(* IEC 61131-3 sources: JingjiangArm/moonboxpro_arm_8.4/Application/Application/任务列表/CommTask/COMM_DIAMONDS/Input_Output (part 3) *)

	i_pstStSysParam^.astStGrpParam_Save[iGrp].rAdjVal_PerTime_Fine			:=	i_pstStParam_Diamonds_WrRd^.arAdjVal_PerTime_Fine[iGrp]   		 	;											(*手动细调调整量*)
	i_pstStSysParam^.astStGrpParam_Save[iGrp].rAdjVal_PerTime_Coarse		:=	i_pstStParam_Diamonds_WrRd^.arAdjVal_PerTime_Coarse[iGrp] 		 	;										(*手动粗调调整量*)
	i_pstStSysParam^.astStGrpParam_Save[iGrp].rVel_HorzdAdj					:=	i_pstStParam_Diamonds_WrRd^.arVel_HorzAdjust[iGrp]        		 	;													(*横向调整速度*)
	i_pstStSysParam^.astStGrpParam_Save[iGrp].rVel_HorzPreRegister			:=	i_pstStParam_Diamonds_WrRd^.arVel_HorzPreRegister[iGrp]   		 	;											(*横向预套准速度*)
	i_pstStSysParam^.astStGrpParam_Save[iGrp].uiNum_If						:=	i_pstStParam_Diamonds_WrRd^.auiNum_If[iGrp]               		 	;														(*放牵减速比-电机侧*)
	i_pstStSysParam^.astStGrpParam_Save[iGrp].uiDen_If						:=	i_pstStParam_Diamonds_WrRd^.auiDen_If[iGrp]               		 	;														(*放牵减速比-传动侧*)
	i_pstStSysParam^.astStGrpParam_Save[iGrp].uiNum_Of						:=	i_pstStParam_Diamonds_WrRd^.auiNum_Of[iGrp]               		 	;														(*收牵减速比-电机侧*)
	i_pstStSysParam^.astStGrpParam_Save[iGrp].uiDen_Of						:=	i_pstStParam_Diamonds_WrRd^.auiDen_Of[iGrp]               		 	;														(*收牵减速比-传动侧*)
	i_pstStSysParam^.astStGrpParam_Save[iGrp].uiNum_Uw						:=	i_pstStParam_Diamonds_WrRd^.auiNum_Uw[iGrp]               		 	;														(*放料减速比-电机侧*)
	i_pstStSysParam^.astStGrpParam_Save[iGrp].uiDen_Uw						:=	i_pstStParam_Diamonds_WrRd^.auiDen_Uw[iGrp]               		 	;														(*放料减速比-传动侧*)
	i_pstStSysParam^.astStGrpParam_Save[iGrp].uiNum_Rw						:=	i_pstStParam_Diamonds_WrRd^.auiNum_Rw[iGrp]               		 	;														(*收料减速比-电机侧*)
	i_pstStSysParam^.astStGrpParam_Save[iGrp].uiDen_Rw						:=	i_pstStParam_Diamonds_WrRd^.auiDen_Rw[iGrp]               		 	;														(*收料减速比-传动侧*)
	i_pstStSysParam^.astStGrpParam_Save[iGrp].uiNum_PrnRoller				:=	i_pstStParam_Diamonds_WrRd^.auiNum_Pu[iGrp]               		 	;												(*色组减速比-电机侧*)
	i_pstStSysParam^.astStGrpParam_Save[iGrp].uiDen_PrnRoller				:=	i_pstStParam_Diamonds_WrRd^.auiDen_Pu[iGrp]               		 	;												(*色组减速比-传动侧*)
	(*待补充-开始|2025.08.07.202603*)
(*	i_pstStSysParam^.astStGrpParam_Save[iGrp].wOutput_IOtestDO_Main[1]		:=	i_pstStParam_Diamonds_WrRd^.awOutput_IOtestDO_Main[iGrp][1]		 	;										(*主面板IO测试输出*)
	i_pstStSysParam^.astStGrpParam_Save[iGrp].wOutput_IOtestDO_Main[2]		:=	i_pstStParam_Diamonds_WrRd^.awOutput_IOtestDO_Main[iGrp][2]		 	;										(*主面板IO测试输出*)
	i_pstStSysParam^.astStGrpParam_Save[iGrp].wOutput_IOtestDO_Main[3]		:=	i_pstStParam_Diamonds_WrRd^.awOutput_IOtestDO_Main[iGrp][3]		 	;										(*主面板IO测试输出*)
	i_pstStSysParam^.astStGrpParam_Save[iGrp].wOutput_IOtestDO_Main[4]		:=	i_pstStParam_Diamonds_WrRd^.awOutput_IOtestDO_Main[iGrp][4]		 	;										(*主面板IO测试输出*)
	i_pstStSysParam^.astStGrpParam_Save[iGrp].wOutput_IOtestDO_Main[5]		:=	i_pstStParam_Diamonds_WrRd^.awOutput_IOtestDO_Main[iGrp][5]		 	;										(*主面板IO测试输出*)
	i_pstStSysParam^.astStGrpParam_Save[iGrp].wOutput_IOtestDO_Main[6]		:=	i_pstStParam_Diamonds_WrRd^.awOutput_IOtestDO_Main[iGrp][6]		 	;										(*主面板IO测试输出*)
	i_pstStSysParam^.astStGrpParam_Save[iGrp].wOutput_IOtestDO_Main[7]		:=	i_pstStParam_Diamonds_WrRd^.awOutput_IOtestDO_Main[iGrp][7]		 	;										(*主面板IO测试输出*)
	i_pstStSysParam^.astStGrpParam_Save[iGrp].wOutput_IOtestDO_Main[8]		:=	i_pstStParam_Diamonds_WrRd^.awOutput_IOtestDO_Main[iGrp][8]		 	;										(*主面板IO测试输出*)

	i_pstStSysParam^.astStGrpParam_Save[iGrp].wOutput_IOtestAO_Main[1]		:=	i_pstStParam_Diamonds_WrRd^.awOutput_IOtestAO_Main[iGrp][1]		 	;									(*主面板IO测试输出*)
	i_pstStSysParam^.astStGrpParam_Save[iGrp].wOutput_IOtestAO_Main[2]		:=	i_pstStParam_Diamonds_WrRd^.awOutput_IOtestAO_Main[iGrp][2]		 	;									(*主面板IO测试输出*)
	i_pstStSysParam^.astStGrpParam_Save[iGrp].wOutput_IOtestAO_Main[3]		:=	i_pstStParam_Diamonds_WrRd^.awOutput_IOtestAO_Main[iGrp][3]		 	;									(*主面板IO测试输出*)
	i_pstStSysParam^.astStGrpParam_Save[iGrp].wOutput_IOtestAO_Main[4]		:=	i_pstStParam_Diamonds_WrRd^.awOutput_IOtestAO_Main[iGrp][4]		 	;									(*主面板IO测试输出*)
	i_pstStSysParam^.astStGrpParam_Save[iGrp].wOutput_IOtestAO_Main[5]		:=	i_pstStParam_Diamonds_WrRd^.awOutput_IOtestAO_Main[iGrp][5]		 	;									(*主面板IO测试输出*)
	i_pstStSysParam^.astStGrpParam_Save[iGrp].wOutput_IOtestAO_Main[6]		:=	i_pstStParam_Diamonds_WrRd^.awOutput_IOtestAO_Main[iGrp][6]		 	;									(*主面板IO测试输出*)
	i_pstStSysParam^.astStGrpParam_Save[iGrp].wOutput_IOtestAO_Main[7]		:=	i_pstStParam_Diamonds_WrRd^.awOutput_IOtestAO_Main[iGrp][7]		 	;									(*主面板IO测试输出*)
	i_pstStSysParam^.astStGrpParam_Save[iGrp].wOutput_IOtestAO_Main[8]		:=	i_pstStParam_Diamonds_WrRd^.awOutput_IOtestAO_Main[iGrp][8]		 	;									(*主面板IO测试输出*)
	i_pstStSysParam^.astStGrpParam_Save[iGrp].wOutput_IOtestAO_Main[9]		:=	i_pstStParam_Diamonds_WrRd^.awOutput_IOtestAO_Main[iGrp][9]		 	;									(*主面板IO测试输出*)
	i_pstStSysParam^.astStGrpParam_Save[iGrp].wOutput_IOtestAO_Main[10]		:=	i_pstStParam_Diamonds_WrRd^.awOutput_IOtestAO_Main[iGrp][10]	 	;										(*主面板IO测试输出*)
	i_pstStSysParam^.astStGrpParam_Save[iGrp].wOutput_IOtestAO_Main[11]		:=	i_pstStParam_Diamonds_WrRd^.awOutput_IOtestAO_Main[iGrp][11]	 	;										(*主面板IO测试输出*)
	i_pstStSysParam^.astStGrpParam_Save[iGrp].wOutput_IOtestAO_Main[12]		:=	i_pstStParam_Diamonds_WrRd^.awOutput_IOtestAO_Main[iGrp][12]	 	;										(*主面板IO测试输出*)
	i_pstStSysParam^.astStGrpParam_Save[iGrp].wOutput_IOtestAO_Main[13]		:=	i_pstStParam_Diamonds_WrRd^.awOutput_IOtestAO_Main[iGrp][13]	 	;										(*主面板IO测试输出*)
	i_pstStSysParam^.astStGrpParam_Save[iGrp].wOutput_IOtestAO_Main[14]		:=	i_pstStParam_Diamonds_WrRd^.awOutput_IOtestAO_Main[iGrp][14]	 	;										(*主面板IO测试输出*)
	i_pstStSysParam^.astStGrpParam_Save[iGrp].wOutput_IOtestAO_Main[15]		:=	i_pstStParam_Diamonds_WrRd^.awOutput_IOtestAO_Main[iGrp][15]	 	;										(*主面板IO测试输出*)
	i_pstStSysParam^.astStGrpParam_Save[iGrp].wOutput_IOtestAO_Main[16]		:=	i_pstStParam_Diamonds_WrRd^.awOutput_IOtestAO_Main[iGrp][16]	 	;										(*主面板IO测试输出*)
*)	(*待补充-结束|2025.08.07.202615*)

	i_pstStSysParam^.astStGrpParam_Save[iGrp].uiPreStopDelayTime_ms		:= 	i_pstStParam_Diamonds_WrRd^.auiPreStopDelayTime_ms[iGrp]    	;
	i_pstStSysParam^.astStGrpParam_Save[iGrp].rVel_Tar_9905				:= 	i_pstStParam_Diamonds_WrRd^.arVel_Tar_9905[iGrp]            	;
	i_pstStSysParam^.astStGrpParam_UnSave[iGrp].iAxisId_StepTest_V		:= 	i_pstStParam_Diamonds_WrRd^.aiAxisId_StepTest_V[iGrp]       	;
	i_pstStSysParam^.astStGrpParam_UnSave[iGrp].iInterval_StepTest12		:= 	i_pstStParam_Diamonds_WrRd^.aiInterval_StepTest12[iGrp]     	;
	i_pstStSysParam^.astStGrpParam_Save[iGrp].iMicron_StepTest1_V		:= 	i_pstStParam_Diamonds_WrRd^.aiMicron_StepTest1_V[iGrp]      	;
	i_pstStSysParam^.astStGrpParam_Save[iGrp].iMicron_StepTest2_V		:= 	i_pstStParam_Diamonds_WrRd^.aiMicron_StepTest2_V[iGrp]      	;
	i_pstStSysParam^.astStGrpParam_Save[iGrp].byKalmanFilterType_Rw		:= 	i_pstStParam_Diamonds_WrRd^.abyKalmanFilterType_Rw[iGrp]    	;
	IF i_pstStParam_Diamonds_WrRd^.abyStructParanInitEn_Rw[iGrp]<>0 THEN
		i_pstStSysParam^.astStGrpParam_Save[iGrp].byStructParanInitEn_Rw 	:= 	i_pstStParam_Diamonds_WrRd^.abyStructParanInitEn_Rw[iGrp]   	;
	END_IF
	i_pstStSysParam^.astStGrpParam_Save[iGrp].rR_K_MinBeat_Rw	    	:= 	i_pstStParam_Diamonds_WrRd^.arR_K_MinBeat_Rw[iGrp]          	;
	i_pstStSysParam^.astStGrpParam_Save[iGrp].iN_MinBeat_Rw	        	:= 	i_pstStParam_Diamonds_WrRd^.aiN_MinBeat_Rw[iGrp]            	;
	i_pstStSysParam^.astStGrpParam_Save[iGrp].rR_K_LQR_Rw	        	:= 	i_pstStParam_Diamonds_WrRd^.arR_K_LQR_Rw[iGrp]              	;

	i_pstStSysParam^.astStGrpParam_Save[iGrp].rN_LQR_Rw	            		:= i_pstStParam_Diamonds_WrRd^.arN_LQR_Rw[iGrp]	               		;
	i_pstStSysParam^.astStGrpParam_Save[iGrp].rKc_Rw	            		:= i_pstStParam_Diamonds_WrRd^.arKc_Rw[iGrp]	                   	;
	i_pstStSysParam^.astStGrpParam_Save[iGrp].rKc_Rw_AccDec	        		:= i_pstStParam_Diamonds_WrRd^.arKc_Rw_AccDec[iGrp]	           		;
	i_pstStSysParam^.astStGrpParam_Save[iGrp].rWc_LowPass_Diam_Rw			:= i_pstStParam_Diamonds_WrRd^.arWc_LowPass_Diam_Rw[iGrp]	   		;
	i_pstStSysParam^.astStGrpParam_Save[iGrp].byKalmanFilterType_Uw 		:= i_pstStParam_Diamonds_WrRd^.abyKalmanFilterType_Uw[iGrp] 	   	;
	IF i_pstStParam_Diamonds_WrRd^.abyStructParanInitEn_Uw[iGrp]<>0 THEN
		i_pstStSysParam^.astStGrpParam_Save[iGrp].byStructParanInitEn_Uw		:= i_pstStParam_Diamonds_WrRd^.abyStructParanInitEn_Uw[iGrp]	   	;
	END_IF
	SysMemCpy(
		ADR(i_pstStSysParam^.astStGrpParam_Save[iGrp].stModelParam_Uw),
		ADR(i_pstStParam_Diamonds_WrRd^.astModelParam_Uw[iGrp]),
		SIZEOF(i_pstStSysParam^.astStGrpParam_Save[iGrp].stModelParam_Uw));
	SysMemCpy(
		ADR(i_pstStSysParam^.astStGrpParam_Save[iGrp].stInvariant_Parameters_Uw),
		ADR(i_pstStParam_Diamonds_WrRd^.astInvariant_Parameters_Uw[iGrp]),
		SIZEOF(i_pstStSysParam^.astStGrpParam_Save[iGrp].stInvariant_Parameters_Uw));
	SysMemCpy(
		ADR(i_pstStSysParam^.astStGrpParam_Save[iGrp].stPI_Parameters_Uw),
		ADR(i_pstStParam_Diamonds_WrRd^.astPI_Parameters_Uw[iGrp]),
		SIZEOF(i_pstStSysParam^.astStGrpParam_Save[iGrp].stPI_Parameters_Uw));
	SysMemCpy(
		ADR(i_pstStSysParam^.astStGrpParam_Save[iGrp].stPI_Parameters_Uw_AccDec),
		ADR(i_pstStParam_Diamonds_WrRd^.astPI_Parameters_Uw_AccDec[iGrp]),
		SIZEOF(i_pstStSysParam^.astStGrpParam_Save[iGrp].stPI_Parameters_Uw_AccDec));

	SysMemCpy(
		ADR(i_pstStSysParam^.astStGrpParam_Save[iGrp].stModelParam_Rw),
		ADR(i_pstStParam_Diamonds_WrRd^.astModelParam_Rw[iGrp]),
		SIZEOF(i_pstStSysParam^.astStGrpParam_Save[iGrp].stModelParam_Rw));
	SysMemCpy(
		ADR(i_pstStSysParam^.astStGrpParam_Save[iGrp].stInvariant_Parameters_Rw),
		ADR(i_pstStParam_Diamonds_WrRd^.astInvariant_Parameters_Rw[iGrp]),
		SIZEOF(i_pstStSysParam^.astStGrpParam_Save[iGrp].stInvariant_Parameters_Rw));
	SysMemCpy(
		ADR(i_pstStSysParam^.astStGrpParam_Save[iGrp].stPI_Parameters_Rw),
		ADR(i_pstStParam_Diamonds_WrRd^.astPI_Parameters_Rw[iGrp]),
		SIZEOF(i_pstStSysParam^.astStGrpParam_Save[iGrp].stPI_Parameters_Rw));
	SysMemCpy(
		ADR(i_pstStSysParam^.astStGrpParam_Save[iGrp].stPI_Parameters_Rw_AccDec),
		ADR(i_pstStParam_Diamonds_WrRd^.astPI_Parameters_Rw_AccDec[iGrp]),
		SIZEOF(i_pstStSysParam^.astStGrpParam_Save[iGrp].stPI_Parameters_Rw_AccDec));

	i_pstStSysParam^.astStGrpParam_Save[iGrp].rR_K_MinBeat_Uw    			:= i_pstStParam_Diamonds_WrRd^.arR_K_MinBeat_Uw[iGrp]    			;
	i_pstStSysParam^.astStGrpParam_Save[iGrp].iN_MinBeat_Uw      			:= i_pstStParam_Diamonds_WrRd^.aiN_MinBeat_Uw[iGrp]      			;
	i_pstStSysParam^.astStGrpParam_Save[iGrp].rR_K_LQR_Uw        			:= i_pstStParam_Diamonds_WrRd^.arR_K_LQR_Uw[iGrp]        			;
	i_pstStSysParam^.astStGrpParam_Save[iGrp].rN_LQR_Uw          			:= i_pstStParam_Diamonds_WrRd^.arN_LQR_Uw[iGrp]          			;
	i_pstStSysParam^.astStGrpParam_Save[iGrp].rKc_Uw             			:= i_pstStParam_Diamonds_WrRd^.arKc_Uw[iGrp]             			;
	i_pstStSysParam^.astStGrpParam_Save[iGrp].rKc_Uw_AccDec      			:= i_pstStParam_Diamonds_WrRd^.arKc_Uw_AccDec[iGrp]      			;
	i_pstStSysParam^.astStGrpParam_Save[iGrp].rWc_LowPass_Diam_Uw			:= i_pstStParam_Diamonds_WrRd^.arWc_LowPass_Diam_Uw[iGrp]			;

	i_pstStSysParam^.astStGrpParam_Save[iGrp].rWn_Uw         				:= i_pstStParam_Diamonds_WrRd^.arWn_Uw[iGrp]         	      		;
	i_pstStSysParam^.astStGrpParam_Save[iGrp].rBw_Uw         				:= i_pstStParam_Diamonds_WrRd^.arBw_Uw[iGrp]         	      		;
	i_pstStSysParam^.astStGrpParam_Save[iGrp].rDp_Uw         				:= i_pstStParam_Diamonds_WrRd^.arDp_Uw[iGrp]         	      		;
	i_pstStSysParam^.astStGrpParam_Save[iGrp].iWorkMode_Pid					:= i_pstStParam_Diamonds_WrRd^.aiWorkMode_Pid[iGrp]		  			;
	i_pstStSysParam^.astStGrpParam_Save[iGrp].rFilmLenth_InUnit  			:= i_pstStParam_Diamonds_WrRd^.arFilmLenth_InUnit[iGrp]	   			;

	(*增加裁切时间集处理2025.9.11.193948*)
	//2026.05.20.214715 替换为直接赋值 by liu.yt
	i_pstStSysParam^.astStGrpParam_UnSave[iGrp].stStTimeSet_DnCut_UpCut_Uw_Hmi:=i_pstStParam_Diamonds_WrRd^.astStTimeSet_DnCut_UpCut_Uw_Hmi[iGrp];
	//2026.05.21.085510 补充收料
	i_pstStSysParam^.astStGrpParam_UnSave[iGrp].stStTimeSet_DnCut_UpCut_RW_Hmi:=i_pstStParam_Diamonds_WrRd^.astStTimeSet_DnCut_UpCut_Rw_Hmi[iGrp];

	i_pstStSysParam^.astStGrpParam_Save[iGrp].byAIType_Uw:= i_pstStParam_Diamonds_WrRd^.abyAIType_Uw[iGrp];
	i_pstStSysParam^.astStGrpParam_Save[iGrp].byAIType_Rw:= i_pstStParam_Diamonds_WrRd^.abyAIType_Rw[iGrp];
	i_pstStSysParam^.astStGrpParam_Save[iGrp].byAIType_If:= i_pstStParam_Diamonds_WrRd^.abyAIType_If[iGrp];
	i_pstStSysParam^.astStGrpParam_Save[iGrp].byAIType_Of:= i_pstStParam_Diamonds_WrRd^.abyAIType_Of[iGrp];
(*2025.10.24.134439||增加变量*)
	i_pstStSysParam^.astStGrpParam_Save[iGrp].byAlarmHold_PreCut_Uw:= i_pstStParam_Diamonds_WrRd^.abyAlarmHold_PreCut_Uw[iGrp];
	i_pstStSysParam^.astStGrpParam_Save[iGrp].byFilmType:= i_pstStParam_Diamonds_WrRd^.abyFilmType[iGrp];
	i_pstStSysParam^.astStGrpParam_Save[iGrp].uiUseTime_Diam_Min_Uw:= i_pstStParam_Diamonds_WrRd^.auiUseTime_Diam_Min_Uw[iGrp];
	i_pstStSysParam^.astStGrpParam_Save[iGrp].uiUseTime_Diam_Min_Rw:= i_pstStParam_Diamonds_WrRd^.auiUseTime_Diam_Min_Rw[iGrp];

(*2025.11.5.154653*)
	i_pstStSysParam^.astStGrpParam_Save[iGrp].iUpperFreq_InkRoller:= i_pstStParam_Diamonds_WrRd^.aiUpperFreq_InkRoller[iGrp];
	i_pstStSysParam^.astStGrpParam_Save[iGrp].iVelSa_InkRollerRun:= i_pstStParam_Diamonds_WrRd^.aiVelSa_InkRollerRun[iGrp];
	i_pstStSysParam^.astStGrpParam_Save[iGrp].iFrq_InkRollerMin:= i_pstStParam_Diamonds_WrRd^.aiFrq_InkRollerMin[iGrp];
	i_pstStSysParam^.astStGrpParam_Save[iGrp].iFrq_InkRollerMax:= i_pstStParam_Diamonds_WrRd^.aiFrq_InkRollerMax[iGrp];
	i_pstStSysParam^.astStGrpParam_Save[iGrp].iVel_InkRollerMin:= i_pstStParam_Diamonds_WrRd^.aiVel_InkRollerMin[iGrp];
	i_pstStSysParam^.astStGrpParam_Save[iGrp].iVel_InkRollerMax:= i_pstStParam_Diamonds_WrRd^.aiVel_InkRollerMax[iGrp];
	i_pstStSysParam^.astStGrpParam_UnSave[iGrp].byPseudoRandomId:= i_pstStParam_Diamonds_WrRd^.abyPseudoRandomId[iGrp];
	i_pstStSysParam^.astStGrpParam_Save[iGrp].rHz_PreHotAir_ManuallySet:= i_pstStParam_Diamonds_WrRd^.arHz_PreHotAir_ManuallySet[iGrp];
	i_pstStSysParam^.astStGrpParam_Save[iGrp].rSV_PreHeating:= i_pstStParam_Diamonds_WrRd^.arSV_PreHeating[iGrp];
	i_pstStSysParam^.astStGrpParam_Save[iGrp].rHz_Scraper_ManuallySet:= i_pstStParam_Diamonds_WrRd^.arHz_Scraper_ManuallySet[iGrp];
	i_pstStSysParam^.astStGrpParam_Save[iGrp].rCoeff_Scraper_Auto:= i_pstStParam_Diamonds_WrRd^.arCoeff_Scraper_Auto[iGrp];
	i_pstStSysParam^.astStGrpParam_Save[iGrp].rHz_InkRoller_ManuallySet:= i_pstStParam_Diamonds_WrRd^.arHz_InkRoller_ManuallySet[iGrp];
	i_pstStSysParam^.astStGrpParam_Save[iGrp].rCoeff_InkRoller:= i_pstStParam_Diamonds_WrRd^.arCoeff_InkRoller_Auto[iGrp];
//2026.1.6.095943增加一些变量
	i_pstStSysParam^.astStGrpParam_Save[iGrp].rLength_Band_Confirm:= i_pstStParam_Diamonds_WrRd^.arLength_Band_Confirm[iGrp];
	i_pstStSysParam^.astStGrpParam_Save[iGrp].rPressure_Tar:= i_pstStParam_Diamonds_WrRd^.arPressure_Tar[iGrp];
// 	xSwitch_TensionAdjust_QH					: BIT;
// 	xSwitch_PrnLenAdj_Follow_QH					: BIT;
	i_pstStSysParam^.stStSysParam_Save.dwCtlSwitchRef.3:= i_pstStParam_Diamonds_WrRd^.astBitStWrRd_Switch_Grp[iGrp].xSwitch_TensionAdjust_QH;
	i_pstStSysParam^.stStSysParam_Save.dwCtlSwitchRef.2:= i_pstStParam_Diamonds_WrRd^.astBitStWrRd_Switch_Grp[iGrp].xSwitch_PrnLenAdj_Follow_QH;

	//2026.2.2.165944||新增界面的一些内容|Niu/j
	i_pstStSysParam^.astStGrpParam_Save[iGrp].rScrewPitch_PrnRoller_Pressure:=
					i_pstStParam_Diamonds_WrRd^.arScrewPitch_PrnRoller_Pressure[iGrp];
	i_pstStSysParam^.astStGrpParam_Save[iGrp].uiNum_PrnRoller_Pressure:=
					i_pstStParam_Diamonds_WrRd^.auiNum_PrnRoller_Pressure[iGrp];
	i_pstStSysParam^.astStGrpParam_Save[iGrp].uiDen_PrnRoller_Pressure:=
					i_pstStParam_Diamonds_WrRd^.auiDen_PrnRoller_Pressure[iGrp];

	i_pstStSysParam^.astStGrpParam_Save[iGrp].rScrewPitch_NetRoller_Pressure:=
					i_pstStParam_Diamonds_WrRd^.arScrewPitch_NetRoller_Pressure[iGrp];
	i_pstStSysParam^.astStGrpParam_Save[iGrp].uiNum_NetRoller_Pressure:=
					i_pstStParam_Diamonds_WrRd^.auiNum_NetRoller_Pressure[iGrp];
	i_pstStSysParam^.astStGrpParam_Save[iGrp].uiDen_NetRoller_Pressure:=
					i_pstStParam_Diamonds_WrRd^.auiDen_NetRoller_Pressure[iGrp];

	i_pstStSysParam^.astStGrpParam_Save[iGrp].rScrewPitch_StrRoller_Pressure:=
					i_pstStParam_Diamonds_WrRd^.arScrewPitch_StrRoller_Pressure[iGrp];
	i_pstStSysParam^.astStGrpParam_Save[iGrp].uiNum_StrRoller_Pressure:=
					i_pstStParam_Diamonds_WrRd^.auiNum_StrRoller_Pressure[iGrp];
	i_pstStSysParam^.astStGrpParam_Save[iGrp].uiDen_StrRoller_Pressure:=
					i_pstStParam_Diamonds_WrRd^.auiDen_StrRoller_Pressure[iGrp];

	i_pstStSysParam^.astStGrpParam_Save[iGrp].rScrewPitch_Horz:=
					i_pstStParam_Diamonds_WrRd^.arScrewPitch_Horz[iGrp];
	i_pstStSysParam^.astStGrpParam_Save[iGrp].uiNum_Horz:=
					i_pstStParam_Diamonds_WrRd^.auiNum_Horz[iGrp];
	i_pstStSysParam^.astStGrpParam_Save[iGrp].uiDen_Horz:=
					i_pstStParam_Diamonds_WrRd^.auiDen_Horz[iGrp];

	i_pstStSysParam^.astStRSV_GrpParam_Save[iGrp].rVel_UVstartVel:= i_pstStParam_Diamonds_WrRd^.arVel_UVstartVel[iGrp];

	//2026.02.28.144731 | + | 上下裁切换
	i_pstStSysParam^.astStGrpParam_Save[iGrp].xSwitch_Change_CutterOnTop_HMI_Uw:=i_pstStParam_Diamonds_WrRd^.astBitStWrRd_Switch_Grp[iGrp].xSwitch_Change_CutterOnTop_HMI_Uw;(*上下裁切换*)
	i_pstStSysParam^.astStGrpParam_Save[iGrp].xSwitch_Change_CutterOnTop_HMI_Rw:=i_pstStParam_Diamonds_WrRd^.astBitStWrRd_Switch_Grp[iGrp].xSwitch_Change_CutterOnTop_HMI_Rw;(*上下裁切换*)

	//2026.03.11.100402 | + | 使用Bit22作为压力电机自动合压开关
	i_pstStSysParam^.astStGrpParam_Save[iGrp].wCtl_Pressure_Up_Dn.0:=i_pstStParam_Diamonds_WrRd^.astBitStWrRd_Switch_Grp[iGrp].xSwitch_PressureAuto_Up_Dn;

	//2026.03.11.114928 | + | 使用Bit24作为停机维持使能的开关
	i_pstStSysParam^.astStGrpParam_Save[iGrp].dwExtBitCtlFlag.21 :=i_pstStParam_Diamonds_WrRd^.astBitStWrRd_Switch_Grp[iGrp].xSwitch_KeepServoOn;

	//2026.02.25.100358 | + | 使用Bit23作为控制天枢存储数据的开关
	i_pstStSysParam^.astStGrpParam_Save[iGrp].dwExtBitCtlFlag.22 :=i_pstStParam_Diamonds_WrRd^.astBitStWrRd_Switch_Grp[iGrp].xSwitch_SaveData_GNS;

	//2026.03.27.175514 | + | 给超旭同步秦华的金刚清除报警功能    2026.1.27.141112 | + | 增加清除报警的功能
	IF 	i_pstStParam_Diamonds_WrRd^.astBitStWrRd_Switch_Grp[iGrp].xSwitch_ClearSysAlarm THEN
		i_pstStParam_Diamonds_WrRd^.astBitStWrRd_Switch_Grp[iGrp].xSwitch_ClearSysAlarm := FALSE;
		g_xClrAlr_HMI := TRUE;
	END_IF
	//2026.04.01.165429 增加总匀墨 Hou.N
	i_pstStSysParam^.astStRSV_GrpParam_UnSave[iGrp].xSwitch_GrpInkEn :=i_pstStParam_Diamonds_WrRd^.astBitStWrRd_Switch_Grp[iGrp].xSwitch_GrpInkEn;
	IF i_pstStParam_Diamonds_WrRd^.astBitStWrRd_Switch_Grp[iGrp].xBtn_ChangeFilmDn_Uw THEN
		i_pstStSysParam^.astStGrpParam_UnSave[iGrp].xCurAxisDia_Uw_Wr:= i_pstStParam_Diamonds_WrRd^.astBitStWrRd_Switch_Grp[iGrp].xBtn_ChangeFilmDn_Uw;
		i_pstStParam_Diamonds_WrRd^.astBitStWrRd_Switch_Grp[iGrp].xBtn_ChangeFilmDn_Uw:= FALSE;
	END_IF
	IF i_pstStParam_Diamonds_WrRd^.astBitStWrRd_Switch_Grp[iGrp].xBtn_ChangeFilmDn_Rw THEN
		i_pstStSysParam^.astStGrpParam_UnSave[iGrp].xCurAxisDia_Rw_Wr:= i_pstStParam_Diamonds_WrRd^.astBitStWrRd_Switch_Grp[iGrp].xBtn_ChangeFilmDn_Rw;
		i_pstStParam_Diamonds_WrRd^.astBitStWrRd_Switch_Grp[iGrp].xBtn_ChangeFilmDn_Rw:= FALSE;
	END_IF
//2026.5.9.172241
	//增加全自动套印相关变量的通讯；2026.4.6.112942|niu.j
	i_pstStSysParam^.astStRSV_GrpParam_UnSave[iGrp].xStartAutoFind:=
		i_pstStParam_Diamonds_WrRd^.astBitStWrRd_Switch_Grp[iGrp].xSwitch_StartAutoFind;
//2026.04.06.141649最终需要放开
	i_pstStSysParam^.astStRSV_GrpParam_Save[iGrp].xSwitch_EnFastPress:=
		i_pstStParam_Diamonds_WrRd^.astBitStWrRd_Switch_Grp[iGrp].xSwitch_EnFastPress;
	i_pstStSysParam^.astStRSV_GrpParam_UnSave[iGrp].xSwitch_SaveRS2file:=
		i_pstStParam_Diamonds_WrRd^.astBitStWrRd_Switch_Grp[iGrp].xSwitch_SaveRS2file;
	i_pstStSysParam^.astStRSV_GrpParam_UnSave[iGrp].xSwitch_RFailure:=
		i_pstStParam_Diamonds_WrRd^.astBitStWrRd_Switch_Grp[iGrp].xSwitch_RFailure;
	i_pstStSysParam^.astStRSV_GrpParam_UnSave[iGrp].xSwitch_FFailure:=
		i_pstStParam_Diamonds_WrRd^.astBitStWrRd_Switch_Grp[iGrp].xSwitch_FFailure;
	i_pstStSysParam^.astStRSV_GrpParam_Save[iGrp].rWidth_Mark_Max:=
			i_pstStParam_Diamonds_WrRd^.arWidth_Mark_Max[iGrp];
	i_pstStSysParam^.astStRSV_GrpParam_Save[iGrp].rWidth_Mark_Min:=
			i_pstStParam_Diamonds_WrRd^.arWidth_Mark_Min[iGrp];
	i_pstStSysParam^.astStRSV_GrpParam_Save[iGrp].rMaxGap:=
			i_pstStParam_Diamonds_WrRd^.arMaxGap[iGrp];
	i_pstStSysParam^.astStRSV_GrpParam_Save[iGrp].bySimilarityThreshold:=
			REAL_TO_BYTE(i_pstStParam_Diamonds_WrRd^.arSimilarityThreshold[iGrp]);
	i_pstStSysParam^.astStRSV_GrpParam_Save[iGrp].byMeanOffset:=
			i_pstStParam_Diamonds_WrRd^.abyMeanOffset[iGrp];
	i_pstStSysParam^.astStRSV_GrpParam_Save[iGrp].bySignalType:=
			i_pstStParam_Diamonds_WrRd^.abySignalType[iGrp];
	i_pstStSysParam^.astStRSV_GrpParam_Save[iGrp].rOuterCoff:=
			i_pstStParam_Diamonds_WrRd^.arOuterCoff[iGrp];
	i_pstStSysParam^.astStRSV_GrpParam_Save[iGrp].rInnerCoff:=
			i_pstStParam_Diamonds_WrRd^.arInnerCoff[iGrp];
	FOR iN:=1 TO 15 BY 1 DO
		IF iN<=2 THEN
			i_pstStSysParam^.astStRSV_GrpParam_Save[iGrp].arFiberMove[iN]:=
						i_pstStParam_Diamonds_WrRd^.arFiberMove[iGrp,iN];
		END_IF
		i_pstStSysParam^.astStRSV_GrpParam_Save[iGrp].arModeMsg[iN]:=
					i_pstStParam_Diamonds_WrRd^.arModeMsg[iGrp,iN];
	END_FOR

	//2026.04.10.110541 增加伪随机pid按钮处理
	i_pstStSysParam^.astStGrpParam_UnSave[iGrp].bySetTestPid_Uw:=i_pstStParam_Diamonds_WrRd^.abySetTestPid_Uw[iGrp];

//2026.4.10.092048增加界面计米清零计数
	IF abyPreCount_ClrPrn[iGrp,1]= i_pstStSysParam^.astStGrpParam_UnSave[iGrp].abyClrPrnLenCount_Rw[1] THEN
		i_pstStSysParam^.astStGrpParam_UnSave[iGrp].abyClrPrnLenCount_Rw[1]:= i_pstStParam_Diamonds_WrRd^.abyClrPrnLenCount[iGrp,1];
	END_IF
	abyPreCount_ClrPrn[iGrp,1]:= i_pstStSysParam^.astStGrpParam_UnSave[iGrp].abyClrPrnLenCount_Rw[1];

	IF abyPreCount_ClrPrn[iGrp,2]= i_pstStSysParam^.astStGrpParam_UnSave[iGrp].abyClrPrnLenCount_Rw[2] THEN
		i_pstStSysParam^.astStGrpParam_UnSave[iGrp].abyClrPrnLenCount_Rw[2]:= i_pstStParam_Diamonds_WrRd^.abyClrPrnLenCount[iGrp,2];
	END_IF
	abyPreCount_ClrPrn[iGrp,2]:= i_pstStSysParam^.astStGrpParam_UnSave[iGrp].abyClrPrnLenCount_Rw[2];

	IF abyPreCount_ClrPrn[iGrp,3]= i_pstStSysParam^.astStGrpParam_UnSave[iGrp].abyClrPrnLenCount_Rw[3] THEN
		i_pstStSysParam^.astStGrpParam_UnSave[iGrp].abyClrPrnLenCount_Rw[3]:= i_pstStParam_Diamonds_WrRd^.abyClrPrnLenCount[iGrp,3];
	END_IF
	abyPreCount_ClrPrn[iGrp,3]:= i_pstStSysParam^.astStGrpParam_UnSave[iGrp].abyClrPrnLenCount_Rw[3];
//增加完成2026.4.10.092101

//2026.5.12.161016增加速度规划方式的通讯
	i_pstStSysParam^.astStGrpParam_Save[iGrp].byAutoAccDecCurve:= i_pstStParam_Diamonds_WrRd^.abyAutoAccDecCurve[iGrp];
	//2026.05.14.151130 新增自动停机、网辊离压速度
    i_pstStSysParam^.astStRSV_GrpParam_Save[iGrp].rRemainDia_stop := i_pstStParam_Diamonds_WrRd^.arRemainDia_stop[iGrp];
    i_pstStSysParam^.astStRSV_GrpParam_Save[iGrp].rMaxErr_GantryTrap := i_pstStParam_Diamonds_WrRd^.arMaxErr_GantryTrap[iGrp];
    i_pstStSysParam^.astStGrpParam_Save[iGrp].rVel_NetReturn := i_pstStParam_Diamonds_WrRd^.arVel_NetReturn[iGrp];
   	i_pstStSysParam^.astStRSV_GrpParam_Save[iGrp].xIsAutoStop :=i_pstStParam_Diamonds_WrRd^.astBitStWrRd_Switch_Grp[iGrp].xSwitch_En_AutoStop;
	//2026.05.15.85606 新增电晕启动速度
	i_pstStSysParam^.astStRSV_GrpParam_Save[iGrp].rVel_CoronaVel:= i_pstStParam_Diamonds_WrRd^.arVel_CoronaVel[iGrp];
	(*2026.05.26.155252+*)
	i_pstStSysParam^.astStGrpParam_UnSave[iGrp].xAutoAccDec_Hmi:=i_pstStParam_Diamonds_WrRd^.astBitStWrRd_Switch_Grp[iGrp].xAutoAccDec_Hmi;

	//2026.05.24.135821 光纤行走部分
	i_pstStSysParam^.astStRSV_GrpParam_Save[iGrp].iFiberMoveVel:=i_pstStParam_Diamonds_WrRd^.aiFiberMoveVel[iGrp];
	i_pstStSysParam^.astStRSV_GrpParam_UnSave[iGrp].rFiberMoveDistance_AllUnit:=i_pstStParam_Diamonds_WrRd^.arFiberMoveDistance_AllUnit[iGrp];
	i_pstStSysParam^.astStRSV_GrpParam_Save[iGrp].byFiberMove_MicroMoveStep:=i_pstStParam_Diamonds_WrRd^.abyFiberMove_MicroMoveStep[iGrp];
	i_pstStSysParam^.astStRSV_GrpParam_UnSave[iGrp].xFiberMove_DebugMode :=i_pstStParam_Diamonds_WrRd^.astBitStWrRd_Switch_Grp[iGrp].xFiberMove_DebugMode;
	i_pstStSysParam^.astStRSV_GrpParam_UnSave[iGrp].xFiberMoveDisRunStart_AllUnit :=i_pstStParam_Diamonds_WrRd^.astBitStWrRd_Switch_Grp[iGrp].xFiberMoveDisRunStart_AllUnit;
	i_pstStSysParam^.astStRSV_GrpParam_Save[iGrp].xUseOnline_FiberMove :=i_pstStParam_Diamonds_WrRd^.astBitStWrRd_Switch_Grp[iGrp].xUseOnline_FiberMove;
	i_pstStSysParam^.astStRSV_GrpParam_UnSave[iGrp].xFiberMoveConfirm_AllUnit :=i_pstStParam_Diamonds_WrRd^.astBitStWrRd_Switch_Grp[iGrp].xFiberMoveConfirm_AllUnit;
	i_pstStSysParam^.astStRSV_GrpParam_UnSave[iGrp].xFiberMovePosCal_ByUnit :=i_pstStParam_Diamonds_WrRd^.astBitStWrRd_Switch_Grp[iGrp].xFiberMovePosCal_ByUnit;
	i_pstStSysParam^.astStRSV_GrpParam_UnSave[iGrp].xFiberMovePosCal_ByOnline :=i_pstStParam_Diamonds_WrRd^.astBitStWrRd_Switch_Grp[iGrp].xFiberMovePosCal_ByOnline;
	i_pstStSysParam^.astStRSV_GrpParam_Save[iGrp].xFiberMove_Negative_AdjustByUnit :=i_pstStParam_Diamonds_WrRd^.astBitStWrRd_Switch_Grp[iGrp].xFiberMove_Negative_AdjustByUnit;
	i_pstStSysParam^.astStRSV_GrpParam_Save[iGrp].xFiberMove_Negative_AdjustByOnline :=i_pstStParam_Diamonds_WrRd^.astBitStWrRd_Switch_Grp[iGrp].xFiberMove_Negative_AdjustByOnline;

//2026.5.15.112026增加卷径检测变量输入
	FOR iK:=1 TO 4 BY 1 DO
		IF arStdVol_Coef_Axis_Hmi_Bak[iGrp,iK]= i_pstStSysParam^.astStGrpParam_UnSave[iGrp].alrStdVol_Coef_Axis_Hmi[iK] THEN
			i_pstStSysParam^.astStGrpParam_UnSave[iGrp].alrStdVol_Coef_Axis_Hmi[iK]:= i_pstStParam_Diamonds_WrRd^.arStdVol_Coef_Axis_Hmi[iGrp,iK];
		END_IF
		arStdVol_Coef_Axis_Hmi_Bak[iGrp,iK]:= i_pstStSysParam^.astStGrpParam_UnSave[iGrp].alrStdVol_Coef_Axis_Hmi[iK];
		IF arStdVol_Diam_Axis_Hmi_Bak[iGrp,iK]= i_pstStSysParam^.astStGrpParam_UnSave[iGrp].alrStdVol_Diam_Axis_Hmi[iK] THEN
			i_pstStSysParam^.astStGrpParam_UnSave[iGrp].alrStdVol_Diam_Axis_Hmi[iK]:=i_pstStParam_Diamonds_WrRd^.arStdVol_Diam_Axis_Hmi[iGrp,iK];
		END_IF
		arStdVol_Diam_Axis_Hmi_Bak[iGrp,iK]:= i_pstStSysParam^.astStGrpParam_UnSave[iGrp].alrStdVol_Diam_Axis_Hmi[iK];
		IF arStdVol_Volt_Axis_Hmi_Bak[iGrp,iK]= i_pstStSysParam^.astStGrpParam_UnSave[iGrp].alrStdVol_Volt_Axis_Hmi[iK] THEN
			i_pstStSysParam^.astStGrpParam_UnSave[iGrp].alrStdVol_Volt_Axis_Hmi[iK]:= i_pstStParam_Diamonds_WrRd^.arStdVol_Volt_Axis_Hmi[iGrp,iK];
		END_IF
		arStdVol_Volt_Axis_Hmi_Bak[iGrp,iK]:= i_pstStSysParam^.astStGrpParam_UnSave[iGrp].alrStdVol_Volt_Axis_Hmi[iK];
	END_FOR
	IF arStdVol_Coef_Axis_Hmi_Bak[iGrp,0]= i_pstStSysParam^.astStGrpParam_UnSave[iGrp].alrStdVol_Coef_Axis_Hmi[0] THEN
		i_pstStSysParam^.astStGrpParam_UnSave[iGrp].alrStdVol_Coef_Axis_Hmi[0]:= i_pstStParam_Diamonds_WrRd^.arStdVol_Coef_Axis_Hmi[iGrp,0];
	END_IF
	arStdVol_Coef_Axis_Hmi_Bak[iGrp,0]:= i_pstStSysParam^.astStGrpParam_UnSave[iGrp].alrStdVol_Coef_Axis_Hmi[0];
END_FOR
(*轴参数|2025.08.07.101610*)
FOR iUnitId:= 1 TO MAX_UNIT_NUM BY 1 DO
	//2026.04.03.115045
	IF axSwitch_AutoAdjust_V_Unit[iUnitId]= i_pstStSysParam^.astStUnitParam_Save[iUnitId].dwFlag_Sts.0 THEN
		i_pstStSysParam^.astStUnitParam_Save[iUnitId].dwFlag_Sts.0 	:=		i_pstStParam_Diamonds_WrRd^.astStWrRd_UnitParam[iUnitId].stBitStWrRd_Switch_Unit.xSwitch_AutoAdjust_V_Unit			 ;			(*整机纵向自动调整开关*)
	END_IF
	axSwitch_AutoAdjust_V_Unit[iUnitId]:= i_pstStSysParam^.astStUnitParam_Save[iUnitId].dwFlag_Sts.0;
	i_pstStSysParam^.astStUnitParam_Save[iUnitId].dwFlag_Sts.1 	:=		i_pstStParam_Diamonds_WrRd^.astStWrRd_UnitParam[iUnitId].stBitStWrRd_Switch_Unit.xSwitch_AutoAdjust_H_Unit			 ;			(*整机纵向自动调整开关*)
	i_pstStSysParam^.astStUnitParam_Save[iUnitId].xEnable_arc 	:=		i_pstStParam_Diamonds_WrRd^.astStWrRd_UnitParam[iUnitId].stBitStWrRd_Switch_Unit.xSwitch_ThisUnitEna ;			(*色组套印开关*)
	i_pstStSysParam^.astStUnitParam_Save[iUnitId].dwFlag_Ctl.0:= i_pstStParam_Diamonds_WrRd^.astStWrRd_UnitParam[iUnitId].stBitStWrRd_Switch_Unit.xSwitch_Horz ;(*横向开关*)
	i_pstStSysParam^.astStUnitParam_Save[iUnitId].dwFlag_Ctl.1:= i_pstStParam_Diamonds_WrRd^.astStWrRd_UnitParam[iUnitId].stBitStWrRd_Switch_Unit.xSwitch_DoorBaseLn	 ;(*门内基线开关*)
	i_pstStSysParam^.astStUnitParam_Save[iUnitId].dwFlag_Ctl.4:= i_pstStParam_Diamonds_WrRd^.astStWrRd_UnitParam[iUnitId].stBitStWrRd_Switch_Unit.xSwitch_AdjRev_V ;(*横向调整反*)
	i_pstStSysParam^.astStUnitParam_Save[iUnitId].dwFlag_Ctl.5:= i_pstStParam_Diamonds_WrRd^.astStWrRd_UnitParam[iUnitId].stBitStWrRd_Switch_Unit.xSwitch_AdjRev_H ;(*横向调整反*)
	i_pstStSysParam^.astStUnitParam_Save[iUnitId].byCouplingMask.2:= i_pstStParam_Diamonds_WrRd^.astStWrRd_UnitParam[iUnitId].stBitStWrRd_Switch_Unit.xSwitch_Transfer_Err ;(*误差传递开关*)
//	i_pstStSysParam^.astStUnitParam_Save[iUnitId].byCouplingMask.0:= i_pstStParam_Diamonds_WrRd^.astStWrRd_UnitParam[iUnitId].stBitStWrRd_Switch_Unit.xSwitch_Transfer_Adj ;(*调整量传递开关*)
(*小信号2025.10.27.141809*)
	i_pstStSysParam^.astStUnitParam_Save[iUnitId].dwFlag_Ctl.13:= i_pstStParam_Diamonds_WrRd^.astStWrRd_UnitParam[iUnitId].stBitStWrRd_Switch_Unit.xSwitch_SmallSignalProcessing_T1;
	i_pstStSysParam^.astStUnitParam_Save[iUnitId].dwFlag_Ctl.14:= i_pstStParam_Diamonds_WrRd^.astStWrRd_UnitParam[iUnitId].stBitStWrRd_Switch_Unit.xSwitch_SmallSignalProcessing_T2;

(*2025.11.12.111108*)
	i_pstStSysParam^.astStUnitParam_Save[iUnitId].xSwitch_ScraperAuto:= i_pstStParam_Diamonds_WrRd^.astStWrRd_UnitParam[iUnitId].stBitStWrRd_Switch_Unit.xSwitch_ScraperAuto ;(*刮刀手自动*)
	i_pstStSysParam^.astStUnitParam_Save[iUnitId].xSwitch_ScraperOn := i_pstStParam_Diamonds_WrRd^.astStWrRd_UnitParam[iUnitId].stBitStWrRd_Switch_Unit.xSwitch_ScraperOn	;(*刮刀开关*)
	i_pstStSysParam^.astStUnitParam_Save[iUnitId].xSwitch_InkRollerAuto:= i_pstStParam_Diamonds_WrRd^.astStWrRd_UnitParam[iUnitId].stBitStWrRd_Switch_Unit.xSwitch_InkRollerAuto ;(*递墨辊手自动*)
	i_pstStSysParam^.astStUnitParam_Save[iUnitId].xSwitch_InkRollerCW := i_pstStParam_Diamonds_WrRd^.astStWrRd_UnitParam[iUnitId].stBitStWrRd_Switch_Unit.xSwitch_InkRollerCW;(*递墨辊正转*)
	i_pstStSysParam^.astStUnitParam_Save[iUnitId].xSwitch_InkRollerCCW:= i_pstStParam_Diamonds_WrRd^.astStWrRd_UnitParam[iUnitId].stBitStWrRd_Switch_Unit.xSwitch_InkRollerCCW ;(*递墨辊反转*)

(*2025.11.5.163824*)
	i_pstStSysParam^.astStUnitParam_Save[iUnitId].xSwitchOn_CoatingPrn:= i_pstStParam_Diamonds_WrRd^.astStWrRd_UnitParam[iUnitId].stBitStWrRd_Switch_Unit.xSwitch_CoatingPrn;(*色组涂布开关*)
	i_pstStSysParam^.astStUnitParam_Save[iUnitId].xReverseAdj_CoatingPrn:= i_pstStParam_Diamonds_WrRd^.astStWrRd_UnitParam[iUnitId].stBitStWrRd_Switch_Unit.xSwitch_CoatingRec;(*涂布调整反向*)
	i_pstStSysParam^.astStUnitParam_Save[iUnitId].xSwitch_HotWindOn:= i_pstStParam_Diamonds_WrRd^.astStWrRd_UnitParam[iUnitId].stBitStWrRd_Switch_Unit.xSwitch_HotWindOn;(*热风开关*)
	i_pstStSysParam^.astStUnitParam_Save[iUnitId].xSwitch_Heating_I:= i_pstStParam_Diamonds_WrRd^.astStWrRd_UnitParam[iUnitId].stBitStWrRd_Switch_Unit.xSwitch_Heating_I;(*加热I档*)
	i_pstStSysParam^.astStUnitParam_Save[iUnitId].xSwitch_Heating_II:= i_pstStParam_Diamonds_WrRd^.astStWrRd_UnitParam[iUnitId].stBitStWrRd_Switch_Unit.xSwitch_Heating_II	;(*加热II档*)
	i_pstStSysParam^.astStUnitParam_Save[iUnitId].xSwitch_Heating_III:= i_pstStParam_Diamonds_WrRd^.astStWrRd_UnitParam[iUnitId].stBitStWrRd_Switch_Unit.xSwitch_Heating_III;(*加热III档*)
	i_pstStSysParam^.astStUnitParam_Save[iUnitId].dwFlag_Ctl.7:= i_pstStParam_Diamonds_WrRd^.astStWrRd_UnitParam[iUnitId].stBitStWrRd_Switch_Unit.xSwitch_AdjRev_O;(*单标记调整反*)
	i_pstStSysParam^.astStUnitParam_Save[iUnitId].dwFlag_Sts.8:= i_pstStParam_Diamonds_WrRd^.astStWrRd_UnitParam[iUnitId].stBitStWrRd_Switch_Unit.xSwitch_Follow_1U_V_Unit;(*纵向跟1色开关*)
	i_pstStSysParam^.astStUnitParam_Save[iUnitId].dwFlag_Sts.9 				:= i_pstStParam_Diamonds_WrRd^.astStWrRd_UnitParam[iUnitId].stBitStWrRd_Switch_Unit.xSwitch_Follow_1U_H_Unit;(*横向跟1色开关*)
	i_pstStSysParam^.astStUnitParam_Save[iUnitId].dwFlag_Ctl.9 				:= i_pstStParam_Diamonds_WrRd^.astStWrRd_UnitParam[iUnitId].stBitStWrRd_Switch_Unit.xSwitch_DualPolarity	;(*双极性开关*)
	i_pstStSysParam^.astStUnitParam_Save[iUnitId].dwFlag_Ctl.8 				:= i_pstStParam_Diamonds_WrRd^.astStWrRd_UnitParam[iUnitId].stBitStWrRd_Switch_Unit.xSwitch_UnitRevPrn		;(*色组反印开关*)
	i_pstStSysParam^.astStUnitParam_Save[iUnitId].dwFlag_Ctl.6 				:= i_pstStParam_Diamonds_WrRd^.astStWrRd_UnitParam[iUnitId].stBitStWrRd_Switch_Unit.xSwitch_DualGate		;(*双波门开关*)
	i_pstStSysParam^.astStUnitParam_Save[iUnitId].byCouplingMask.2 			:= i_pstStParam_Diamonds_WrRd^.astStWrRd_UnitParam[iUnitId].stBitStWrRd_Switch_Unit.xSwitch_Transfer_Err	;(*误差传递开关*)
	i_pstStSysParam^.astStUnitParam_Save[iUnitId].byCouplingMask.0 			:= i_pstStParam_Diamonds_WrRd^.astStWrRd_UnitParam[iUnitId].stBitStWrRd_Switch_Unit.xSwitch_Transfer_Adj	;(*调整量传递开关*)
//2026.5.12.163836增加小信号处理
//小信号 2026.05.11.191235
	i_pstStSysParam^.astStUnitParam_Save[iUnitId].dwFlag_Ctl.13:=i_pstStParam_Diamonds_WrRd^.astStWrRd_UnitParam[iUnitId].stBitStWrRd_Switch_Unit.xSwitch_SmallSignalProcessing_T1	;
	i_pstStSysParam^.astStUnitParam_Save[iUnitId].dwFlag_Ctl.14:=i_pstStParam_Diamonds_WrRd^.astStWrRd_UnitParam[iUnitId].stBitStWrRd_Switch_Unit.xSwitch_SmallSignalProcessing_T2	;

//2026.5.11.172229+反极性值界面修改未赋值
	i_pstStSysParam^.astStUnitParam_Save[iUnitId].dwFlag_Ctl.2 :=i_pstStParam_Diamonds_WrRd^.astStWrRd_UnitParam[iUnitId].stBitStWrRd_Switch_Unit.xSwitch_NegativePolarity_T1_1	;(*第一组波门内T1信号反极性*)
	i_pstStSysParam^.astStUnitParam_Save[iUnitId].dwFlag_Ctl.3 :=i_pstStParam_Diamonds_WrRd^.astStWrRd_UnitParam[iUnitId].stBitStWrRd_Switch_Unit.xSwitch_NegativePolarity_T2_1	;(*第一组波门内T2信号反极性*)
	i_pstStSysParam^.astStUnitParam_Save[iUnitId].dwFlag_Ctl.11:=i_pstStParam_Diamonds_WrRd^.astStWrRd_UnitParam[iUnitId].stBitStWrRd_Switch_Unit.xSwitch_NegativePolarity_T1_2	;(*第二组波门内T1信号反极性*)
	i_pstStSysParam^.astStUnitParam_Save[iUnitId].dwFlag_Ctl.12:=i_pstStParam_Diamonds_WrRd^.astStWrRd_UnitParam[iUnitId].stBitStWrRd_Switch_Unit.xSwitch_NegativePolarity_T2_2	;(*第二组波门内T2信号反极性*)
//2026.5.12.163844

	i_pstStSysParam^.astStUnitParam_Save[iUnitId].xSwitch_HeatingMode_Water := i_pstStParam_Diamonds_WrRd^.astStWrRd_UnitParam[iUnitId].stBitStWrRd_Switch_Unit.xSwitch_Heating_Water	;(*水加热控制开关*)
	i_pstStSysParam^.astStUnitParam_Save[iUnitId].xSwitch_HeatingMode_Ele 	:= i_pstStParam_Diamonds_WrRd^.astStWrRd_UnitParam[iUnitId].stBitStWrRd_Switch_Unit.xSwitch_Heating_Elc	;(*电加热控制开关*)
	i_pstStSysParam^.astStUnitParam_Save[iUnitId].xSwitch_ExhAir 			:= i_pstStParam_Diamonds_WrRd^.astStWrRd_UnitParam[iUnitId].stBitStWrRd_Switch_Unit.xSwitch_ExhAir			;(*色组排风开关*)
	i_pstStSysParam^.astStUnitParam_Save[iUnitId].stStArc_Mol_Param.xCompensateEn_H 	:= i_pstStParam_Diamonds_WrRd^.astStWrRd_UnitParam[iUnitId].stBitStWrRd_Switch_Unit.xCompensateEn_H	;
	i_pstStSysParam^.astStUnitParam_Save[iUnitId].stStArc_Mol_Param.xUseAntiNotch_Arc 	:= i_pstStParam_Diamonds_WrRd^.astStWrRd_UnitParam[iUnitId].stBitStWrRd_Switch_Unit.xUseAntiNotch_Arc  ;
	i_pstStSysParam^.astStUnitParam_Save[iUnitId].stStArc_Mol_Param.xUsePeriodic 		:= i_pstStParam_Diamonds_WrRd^.astStWrRd_UnitParam[iUnitId].stBitStWrRd_Switch_Unit.xUsePeriodic    	;

	i_pstStSysParam^.astStUnitParam_Save[iUnitId].lrGirth_Using_CoatingPrn 			:=	i_pstStParam_Diamonds_WrRd^.astStWrRd_UnitParam[iUnitId].rGirth_Using_CoatingPrn			 ;  		(*涂布周长*)
	i_pstStSysParam^.astStUnitParam_Save[iUnitId].byAdjMode_CoatingPrn 				:=	i_pstStParam_Diamonds_WrRd^.astStWrRd_UnitParam[iUnitId].byBtn_AdjModeSwitch_CoatingPrn		 ;      	(*涂布调整方式切换按钮*)
	i_pstStSysParam^.astStUnitParam_Save[iUnitId].rStep_OfChangeGirth 				:=	i_pstStParam_Diamonds_WrRd^.astStWrRd_UnitParam[iUnitId].rStep_OfChangeGirth				 ;  		(*涂布版轴修改步幅*)
	i_pstStSysParam^.astStUnitParam_Save[iUnitId].rHz_UnitScraper_ManuallySet 		:=	i_pstStParam_Diamonds_WrRd^.astStWrRd_UnitParam[iUnitId].rHz_UnitScraper_ManuallySet		 ;  		(*刮刀手动频率*)
	i_pstStSysParam^.astStUnitParam_Save[iUnitId].rCoeff_UnitScraper_Auto 			:=	i_pstStParam_Diamonds_WrRd^.astStWrRd_UnitParam[iUnitId].rCoeff_UnitScraper_Auto			 ;  		(*刮刀自动系数*)
	i_pstStSysParam^.astStUnitParam_Save[iUnitId].rHz_UnitInkRoller_ManuallySet 	:=	i_pstStParam_Diamonds_WrRd^.astStWrRd_UnitParam[iUnitId].rHz_UnitInkRoller_ManuallySet		 ;			(*递墨辊手动频率*)
	i_pstStSysParam^.astStUnitParam_Save[iUnitId].rCoeff_UnitInkRoller_Auto 		:=	i_pstStParam_Diamonds_WrRd^.astStWrRd_UnitParam[iUnitId].rCoeff_UnitInkRoller_Auto			 ;    		(*递墨辊自动系数*)
	i_pstStSysParam^.astStUnitParam_Save[iUnitId].rHz_UnitHotWind_ManuallySet 		:=	i_pstStParam_Diamonds_WrRd^.astStWrRd_UnitParam[iUnitId].rHz_UnitHotWind_ManuallySet		 ;  		(*热风手动频率*)
	i_pstStSysParam^.astStUnitParam_Save[iUnitId].rSV_UnitTemCtl 					:=	i_pstStParam_Diamonds_WrRd^.astStWrRd_UnitParam[iUnitId].rSV_UnitTemCtl						 ;      	(*加热设定温度*)
	i_pstStSysParam^.astStUnitParam_Save[iUnitId].iGateWidthPhy 					:=	i_pstStParam_Diamonds_WrRd^.astStWrRd_UnitParam[iUnitId].iGateWidthPhy						 ;      	(*波门宽度*)
	i_pstStSysParam^.astStUnitParam_Save[iUnitId].rAlr_V 							:=	i_pstStParam_Diamonds_WrRd^.astStWrRd_UnitParam[iUnitId].rAlarm_V							 ;      	(*纵向报警值*)
	i_pstStSysParam^.astStUnitParam_Save[iUnitId].rAlr_H 							:=	i_pstStParam_Diamonds_WrRd^.astStWrRd_UnitParam[iUnitId].rAlarm_H							 ;      	(*横向报警值*)
	i_pstStSysParam^.astStUnitParam_Save[iUnitId].rAdj_V 							:=	i_pstStParam_Diamonds_WrRd^.astStWrRd_UnitParam[iUnitId].rAdjust_V							 ;      	(*纵向修正量*)
	i_pstStSysParam^.astStUnitParam_Save[iUnitId].rAdj_H 							:=	i_pstStParam_Diamonds_WrRd^.astStWrRd_UnitParam[iUnitId].rAdjust_H							 ;      	(*横向修正量*)
	i_pstStSysParam^.astStUnitParam_Save[iUnitId].rDeadzoneMax_H 					:=	i_pstStParam_Diamonds_WrRd^.astStWrRd_UnitParam[iUnitId].rDeadzoneMax_H						 ;      	(*横向最大不动作区*)
	i_pstStSysParam^.astStUnitParam_Save[iUnitId].rDeadzoneMin_H 					:=	i_pstStParam_Diamonds_WrRd^.astStWrRd_UnitParam[iUnitId].rDeadzoneMin_H						 ;      	(*横向最小不动作区*)
	i_pstStSysParam^.astStUnitParam_Save[iUnitId].iCoefOfCoupling_V 				:=	i_pstStParam_Diamonds_WrRd^.astStWrRd_UnitParam[iUnitId].iCoefOfCoupling_V					 ;      	(*纵向传递2系数*)
	i_pstStSysParam^.astStUnitParam_Save[iUnitId].byAvg_V 							:=	i_pstStParam_Diamonds_WrRd^.astStWrRd_UnitParam[iUnitId].byAverage_V						 ;  		(*纵向平均值*)
	i_pstStSysParam^.astStUnitParam_Save[iUnitId].byAvg_H 							:=	i_pstStParam_Diamonds_WrRd^.astStWrRd_UnitParam[iUnitId].byAverage_H						 ;  		(*横向平均值*)
	(*待补充-开始|2025.08.07.204217*)
	(*待补充-结束|2025.08.07.204230*)
	i_pstStSysParam^.astStUnitParam_Save[iUnitId].uiTimeMs_RollerPressUpKeep 	:= i_pstStParam_Diamonds_WrRd^.astStWrRd_UnitParam[iUnitId].uiTimeMs_RollerPressUpKeep			;       (*压辊双气缸-离压保持时间*)
	i_pstStSysParam^.astStUnitParam_Save[iUnitId].uiNum_PrnRoller 				:= i_pstStParam_Diamonds_WrRd^.astStWrRd_UnitParam[iUnitId].uiAxisNum							;      			(*色组单独减速比分子*)
	i_pstStSysParam^.astStUnitParam_Save[iUnitId].uiDen_PrnRoller 				:= i_pstStParam_Diamonds_WrRd^.astStWrRd_UnitParam[iUnitId].uiAxisDen							;     				(*色组单独减速比分母*)
	i_pstStSysParam^.astStUnitParam_Save[iUnitId].rHz_UnitExhaust_ManuallySet 	:= i_pstStParam_Diamonds_WrRd^.astStWrRd_UnitParam[iUnitId].rHz_UnitExhaust_ManuallySet		;  	(*色组排风设定频率*)
	//9905界面内容
	i_pstStSysParam^.astStUnitParam_Save[iUnitId].rAxisVelPrf_Coeff1 			:= 	i_pstStParam_Diamonds_WrRd^.astStWrRd_UnitParam[iUnitId].rAxisVelPrf_Coeff1						;
	i_pstStSysParam^.astStUnitParam_Save[iUnitId].rAxisVelPrf_Coeff2 			:= 	i_pstStParam_Diamonds_WrRd^.astStWrRd_UnitParam[iUnitId].rAxisVelPrf_Coeff2             		;
	i_pstStSysParam^.astStUnitParam_Save[iUnitId].rAxisVelPrf_Coeff3 			:= 	i_pstStParam_Diamonds_WrRd^.astStWrRd_UnitParam[iUnitId].rAxisVelPrf_Coeff3             		;
	i_pstStSysParam^.astStUnitParam_Save[iUnitId].stStArc_Mol_Param.rMargin_Mag_Arc 				:= 	i_pstStParam_Diamonds_WrRd^.astStWrRd_UnitParam[iUnitId].rMargin_Mag_Arc                		;
//	//2026.05.13.091849+变量替换
	i_pstStSysParam^.astStUnitParam_Save[iUnitId].stStArc_Mol_Param.rKadj_I_Mol 	:= 	i_pstStParam_Diamonds_WrRd^.astStWrRd_UnitParam[iUnitId].rKadj_I_Mol                		;
//	i_pstStSysParam^.astStUnitParam_Save[iUnitId].rMargin_Phi_Arc 				:= 	i_pstStParam_Diamonds_WrRd^.astStWrRd_UnitParam[iUnitId].rMargin_Phi_Arc                		;
//这两个变量放只写区域，不需要双向2026.4.25.142438
//	i_pstStSysParam^.astStUnitParam_Save[iUnitId].rKp_MolCal 					:= 	i_pstStParam_Diamonds_WrRd^.astStWrRd_UnitParam[iUnitId].rKp_MolCal                     		;
//	i_pstStSysParam^.astStUnitParam_Save[iUnitId].rKi_MolCal 					:= 	i_pstStParam_Diamonds_WrRd^.astStWrRd_UnitParam[iUnitId].rKi_MolCal                     		;
//2026.4.25.142452结束
	i_pstStSysParam^.astStUnitParam_Save[iUnitId].rFilmLengthFromPrevPressUnit 	:= 	i_pstStParam_Diamonds_WrRd^.astStWrRd_UnitParam[iUnitId].rFilmLengthFromPrevPressUnit   		;
	i_pstStSysParam^.astStUnitParam_Save[iUnitId].byCompensateValue_Hor 		:= 	i_pstStParam_Diamonds_WrRd^.astStWrRd_UnitParam[iUnitId].byCompensateValue_Hor					;
	i_pstStSysParam^.astStUnitParam_Save[iUnitId].byMaxAddValue_Total_Hor 		:= 	i_pstStParam_Diamonds_WrRd^.astStWrRd_UnitParam[iUnitId].byMaxAddValue_Total_Hor				;
	i_pstStSysParam^.astStUnitParam_Save[iUnitId].rWn_Arc 						:= 	i_pstStParam_Diamonds_WrRd^.astStWrRd_UnitParam[iUnitId].rWn_Arc								;
	i_pstStSysParam^.astStUnitParam_Save[iUnitId].rBw_Arc 						:= 	i_pstStParam_Diamonds_WrRd^.astStWrRd_UnitParam[iUnitId].rBw_Arc								;
	i_pstStSysParam^.astStUnitParam_Save[iUnitId].rDp_Arc 						:= 	i_pstStParam_Diamonds_WrRd^.astStWrRd_UnitParam[iUnitId].rDp_Arc								;
	i_pstStSysParam^.astStUnitParam_Save[iUnitId].rK 							:= 	i_pstStParam_Diamonds_WrRd^.astStWrRd_UnitParam[iUnitId].rK     								;
	i_pstStSysParam^.astStUnitParam_Save[iUnitId].rA2 							:= 	i_pstStParam_Diamonds_WrRd^.astStWrRd_UnitParam[iUnitId].rA2    								;
	i_pstStSysParam^.astStUnitParam_Save[iUnitId].rA1 							:= 	i_pstStParam_Diamonds_WrRd^.astStWrRd_UnitParam[iUnitId].rA1    								;
	i_pstStSysParam^.astStUnitParam_Save[iUnitId].rA0 							:= 	i_pstStParam_Diamonds_WrRd^.astStWrRd_UnitParam[iUnitId].rA0    								;
	i_pstStSysParam^.astStUnitParam_Save[iUnitId].rG_Periodic 					:= 	i_pstStParam_Diamonds_WrRd^.astStWrRd_UnitParam[iUnitId].rG_Periodic  							;
	i_pstStSysParam^.astStUnitParam_Save[iUnitId].rW_Periodic 					:= 	i_pstStParam_Diamonds_WrRd^.astStWrRd_UnitParam[iUnitId].rW_Periodic  							;
	i_pstStSysParam^.astStUnitParam_Save[iUnitId].byCnt_Comm2ARM 				:= 	i_pstStParam_Diamonds_WrRd^.astStWrRd_UnitParam[iUnitId].byCnt_Comm2ARM							;

(*2025.8.25.151756|、niu.j||波门位置*)
(*2025.8.25.151756|、niu.j||波门位置*)
	//2026.04.03.115113
	IF aiGateSa_Pre_GNS[iUnitId]=i_pstStSysParam^.astStUnitParam_Save[iUnitId].iGateSa THEN
		i_pstStSysParam^.astStUnitParam_Save[iUnitId].iGateSa:= i_pstStParam_Diamonds_WrRd^.astStWrRd_UnitParam[iUnitId].iGateSa	;
	END_IF
	aiGateSa_Pre_GNS[iUnitId]:=i_pstStSysParam^.astStUnitParam_Save[iUnitId].iGateSa;
	i_pstStSysParam^.astStUnitParam_Save[iUnitId].iGateSaEx:= i_pstStParam_Diamonds_WrRd^.astStWrRd_UnitParam[iUnitId].iGateSaEx	;
(*2025.9.19.124046*)
	i_pstStSysParam^.astStUnitParam_Save[iUnitId].iMarkArrangeMode:= i_pstStParam_Diamonds_WrRd^.astStWrRd_UnitParam[iUnitId].iMarkArrangeMode;
(*横向手动调整按钮2025.9.20.111304*)
	g_abyHorzManu_HMI[iUnitId].0 := i_pstStParam_Diamonds_WrRd^.astStWrRd_UnitParam[iUnitId].stBitStWrRd_Switch_Unit.xSwitch_HorzMoveLeft_Manu_1;
	g_abyHorzManu_HMI[iUnitId].4 := i_pstStParam_Diamonds_WrRd^.astStWrRd_UnitParam[iUnitId].stBitStWrRd_Switch_Unit.xSwitch_HorzMoveLeft_Manu_2;
	g_abyHorzManu_HMI[iUnitId].1 := i_pstStParam_Diamonds_WrRd^.astStWrRd_UnitParam[iUnitId].stBitStWrRd_Switch_Unit.xSwitch_HorzMoveLeft_Manu_3;
	g_abyHorzManu_HMI[iUnitId].2 := i_pstStParam_Diamonds_WrRd^.astStWrRd_UnitParam[iUnitId].stBitStWrRd_Switch_Unit.xSwitch_HorzMoveRight_Manu_1;
	g_abyHorzManu_HMI[iUnitId].5 := i_pstStParam_Diamonds_WrRd^.astStWrRd_UnitParam[iUnitId].stBitStWrRd_Switch_Unit.xSwitch_HorzMoveRight_Manu_2;
	g_abyHorzManu_HMI[iUnitId].3 := i_pstStParam_Diamonds_WrRd^.astStWrRd_UnitParam[iUnitId].stBitStWrRd_Switch_Unit.xSwitch_HorzMoveRight_Manu_3;

(*2025.11.5.165752*)
	i_pstStSysParam^.astStUnitParam_Save[iUnitId].lrPreReg_Adjust:= i_pstStParam_Diamonds_WrRd^.astStWrRd_UnitParam[iUnitId].rPreReg_Adjust;
	i_pstStSysParam^.astStUnitParam_Save[iUnitId].lrPreReg_ConstVal:= i_pstStParam_Diamonds_WrRd^.astStWrRd_UnitParam[iUnitId].rPreReg_ConstVal;
	i_pstStSysParam^.astStUnitParam_Save[iUnitId].uiTurnOverFilmLenth:= i_pstStParam_Diamonds_WrRd^.astStWrRd_UnitParam[iUnitId].uiTurnOverFilmLenth;
	i_pstStSysParam^.astStUnitParam_UnSave[iUnitId].diPreReg_RepeatVal_H:= i_pstStParam_Diamonds_WrRd^.astStWrRd_UnitParam[iUnitId].diPreReg_RepeatVal_H;
	i_pstStSysParam^.astStUnitParam_UnSave[iUnitId].diPreReg_SetupVal_H:= i_pstStParam_Diamonds_WrRd^.astStWrRd_UnitParam[iUnitId].diPreReg_SetupVal_H;
	i_pstStSysParam^.astStUnitParam_Save[iUnitId].diPreReg_AdjustVal_H:= i_pstStParam_Diamonds_WrRd^.astStWrRd_UnitParam[iUnitId].diPreReg_AdjustVal_H;

	i_pstStSysParam^.astStUnitParam_Save[iUnitId].rGirth_PrnRoller:= i_pstStParam_Diamonds_WrRd^.astStWrRd_UnitParam[iUnitId].rGirth_PrnRoller;
	i_pstStSysParam^.astStUnitParam_Save[iUnitId].byAirInletWindDoorValue:= i_pstStParam_Diamonds_WrRd^.astStWrRd_UnitParam[iUnitId].byAirInletWindDoorValue;
//	i_pstStSysParam^.astStUnitParam_Save[iUnitId].byOvensAirOutWindDoorValue:= i_pstStParam_Diamonds_WrRd^.astStWrRd_UnitParam[iUnitId].byAirInletWindDoorValue;
	i_pstStSysParam^.astStUnitParam_Save[iUnitId].wAirReturnWindDoorValue:= BYTE_TO_WORD(i_pstStParam_Diamonds_WrRd^.astStWrRd_UnitParam[iUnitId].byAirReturnWindDoorValue);
	i_pstStSysParam^.astStUnitParam_Save[iUnitId].wAirExhaustWindDoorValue:= BYTE_TO_WORD(i_pstStParam_Diamonds_WrRd^.astStWrRd_UnitParam[iUnitId].byAirExhaustWindDoorValue);
	i_pstStSysParam^.astStUnitParam_Save[iUnitId].byOvensAirOutWindDoorValue        := i_pstStParam_Diamonds_WrRd^.astStWrRd_UnitParam[iUnitId].byAirInletWindDoorValue;
	i_pstStSysParam^.astStUnitParam_Save[iUnitId].byFakeThreshold_V:= i_pstStParam_Diamonds_WrRd^.astStWrRd_UnitParam[iUnitId].byFakeThreshold_V;
	i_pstStSysParam^.astStUnitParam_Save[iUnitId].byFakeThreshold_H:= i_pstStParam_Diamonds_WrRd^.astStWrRd_UnitParam[iUnitId].byFakeThreshold_H;
	i_pstStSysParam^.astStUnitParam_Save[iUnitId].byAve_v_extra:= i_pstStParam_Diamonds_WrRd^.astStWrRd_UnitParam[iUnitId].byAve_v_extra;

//2026.1.6.095943增加一些变量
	i_pstStSysParam^.astStUnitParam_Save[iUnitId].iBandLengthFilterCnt:= i_pstStParam_Diamonds_WrRd^.astStWrRd_UnitParam[iUnitId].iBandLengthFilterCnt;
 	i_pstStSysParam^.astStUnitParam_UnSave[iUnitId].xAdjBandLen:= i_pstStParam_Diamonds_WrRd^.astStWrRd_UnitParam[iUnitId].stBitStWrRd_Switch_Unit.xSwitch_AdjBandLen;
	//2026.2.2.165944||新增界面的一些内容|Niu/j

	IF i_pstStParam_Diamonds_WrRd^.astStWrRd_UnitParam[iUnitId].adwPressureMotor_Move_MasterHMI[1]<>0 THEN
		i_pstStSysParam^.astStUnitParam_UnSave[iUnitId].adwPressureMotor_Move[1]:=
				i_pstStParam_Diamonds_WrRd^.astStWrRd_UnitParam[iUnitId].adwPressureMotor_Move_MasterHMI[1];
		i_pstStParam_Diamonds_WrRd^.astStWrRd_UnitParam[iUnitId].adwPressureMotor_Move_MasterHMI[1]:= 0;
	END_IF
	IF i_pstStParam_Diamonds_WrRd^.astStWrRd_UnitParam[iUnitId].adwPressureMotor_Move_MasterHMI[2]<>0 THEN
		i_pstStSysParam^.astStUnitParam_UnSave[iUnitId].adwPressureMotor_Move[2]:=
				i_pstStParam_Diamonds_WrRd^.astStWrRd_UnitParam[iUnitId].adwPressureMotor_Move_MasterHMI[2];
		i_pstStParam_Diamonds_WrRd^.astStWrRd_UnitParam[iUnitId].adwPressureMotor_Move_MasterHMI[2]:= 0;
	END_IF
	IF i_pstStParam_Diamonds_WrRd^.astStWrRd_UnitParam[iUnitId].adwPressureMotor_Move_MasterHMI[3]<>0 THEN
		i_pstStSysParam^.astStUnitParam_UnSave[iUnitId].adwPressureMotor_Move[3]:=
				i_pstStParam_Diamonds_WrRd^.astStWrRd_UnitParam[iUnitId].adwPressureMotor_Move_MasterHMI[3];
		i_pstStParam_Diamonds_WrRd^.astStWrRd_UnitParam[iUnitId].adwPressureMotor_Move_MasterHMI[3]:= 0;
	END_IF

	//2026.02.06.194535增加联动和匀墨
	(*变量使用错误@2026.06.02.130846+*)
	i_pstStSysParam^.astStRSV_UnitParam_Save[iUnitId].xSwitch_Linkage :=
							i_pstStParam_Diamonds_WrRd^.astStWrRd_UnitParam[iUnitId].stBitStWrRd_Switch_Unit.xSwitch_Linkage;
	i_pstStSysParam^.astStUnitParam_Save[iUnitId].wSwitchFun.0 :=
							i_pstStSysParam^.astStRSV_UnitParam_Save[iUnitId].xSwitch_Linkage;

	i_pstStSysParam^.astStRSV_UnitParam_UnSave[iUnitId].xSwitch_Inching_Net
				:= i_pstStParam_Diamonds_WrRd^.astStWrRd_UnitParam[iUnitId].stBitStWrRd_Switch_Unit.xSwitch_Ink;

	//2026.04.02.191415  Hou.N 增加横向限位实时位置
	g_axLimit_Left_Wr[iUnitId]:=i_pstStParam_Diamonds_WrRd^.astStWrRd_UnitParam[iUnitId].stBitStWrRd_Switch_Unit.xBtn_ConfirmLimit_Left	 ;(*标定横向左限位*)
    g_axLimit_Right_Wr[iUnitId]:=i_pstStParam_Diamonds_WrRd^.astStWrRd_UnitParam[iUnitId].stBitStWrRd_Switch_Unit.xBtn_ConfirmLimit_Right;(*标定横向右限位*)
    g_axLimit_Left_WrClr[iUnitId]:=i_pstStParam_Diamonds_WrRd^.astStWrRd_UnitParam[iUnitId].stBitStWrRd_Switch_Unit.xBtn_ResetLimit_Left;(*清除横向左限位*)
    g_axLimit_Right_WrClr[iUnitId]:=i_pstStParam_Diamonds_WrRd^.astStWrRd_UnitParam[iUnitId].stBitStWrRd_Switch_Unit.xBtn_ResetLimit_Right ;(*清除横向右限位*)
//2026.5.10.002039
	IF NOT i_pstStSysParam^.astStRSV_UnitParam_UnSave[iUnitId].xBtn_FromHMI_HorMove_G THEN
		i_pstStSysParam^.astStRSV_UnitParam_UnSave[iUnitId].xBtn_FromHMI_HorMove_G:= i_pstStParam_Diamonds_WrRd^.astStWrRd_UnitParam[iUnitId].stBitStWrRd_Switch_Unit.xBtn_MoveLeft_Horz;(*横向左移*)
		i_pstStParam_Diamonds_WrRd^.astStWrRd_UnitParam[iUnitId].stBitStWrRd_Switch_Unit.xBtn_MoveLeft_Horz:= FALSE;
	END_IF
	IF NOT i_pstStSysParam^.astStRSV_UnitParam_UnSave[iUnitId].xBtn_FromHMI_HorMove_M THEN
		i_pstStSysParam^.astStRSV_UnitParam_UnSave[iUnitId].xBtn_FromHMI_HorMove_M:=i_pstStParam_Diamonds_WrRd^.astStWrRd_UnitParam[iUnitId].stBitStWrRd_Switch_Unit.xBtn_MoveRight_Horz ;(*横向右移*)
		i_pstStParam_Diamonds_WrRd^.astStWrRd_UnitParam[iUnitId].stBitStWrRd_Switch_Unit.xBtn_MoveRight_Horz:= FALSE;
	END_IF

//	i_pstStSysParam^.astStUnitParam_UnSave[iUnitId].lrLimit_Left:=
	i_pstStSysParam^.astStRSV_UnitParam_Save[iUnitId].lrLimit_Left:=
				DINT_TO_LREAL(i_pstStParam_Diamonds_WrRd^.astStWrRd_UnitParam[iUnitId].diPos_LimitLeft);
//	i_pstStSysParam^.astStUnitParam_UnSave[iUnitId].lrLimit_Right:=
	i_pstStSysParam^.astStRSV_UnitParam_Save[iUnitId].lrLimit_Right:=
				DINT_TO_LREAL(i_pstStParam_Diamonds_WrRd^.astStWrRd_UnitParam[iUnitId].diPos_LimitRight);
// 	g_alrTrap_EncPos[iUnitId]:=
// 				DINT_TO_LREAL(i_pstStParam_Diamonds_WrRd^.astStWrRd_UnitParam[iUnitId].diPos_Horz);

//增加全自动套印相关变量2026.4.6.130533|2026.5.9.172510
	i_pstStSysParam^.astStRSV_UnitParam_UnSave[iUnitId].xCurManuAdjust:=
				i_pstStParam_Diamonds_WrRd^.astStWrRd_UnitParam[iUnitId].stBitStWrRd_Switch_Unit.xSwitch_CurManuAdjust;
	i_pstStSysParam^.astStRSV_UnitParam_UnSave[iUnitId].xPreCurManuAdjust:=
				i_pstStParam_Diamonds_WrRd^.astStWrRd_UnitParam[iUnitId].stBitStWrRd_Switch_Unit.xSwitch_PreCurManuAdjust;

//2026.05.24.180357 光纤行走
i_pstStSysParam^.astStRSV_UnitParam_Save[iUnitId].rFiberMoveAdjust:=i_pstStParam_Diamonds_WrRd^.astStWrRd_UnitParam[iUnitId].rFiberMoveAdjust;
i_pstStSysParam^.astStRSV_UnitParam_Save[iUnitId].rFiberMoveAdjust_ByOnlie:=i_pstStParam_Diamonds_WrRd^.astStWrRd_UnitParam[iUnitId].rFiberMoveAdjust_ByOnlie;
//2026.5.29.172542增加一些变量
i_pstStSysParam^.astStUnitParam_Save[iUnitId].xSwitch_Coolwind:=
			i_pstStParam_Diamonds_WrRd^.astStWrRd_UnitParam[iUnitId].stBitStWrRd_Switch_Unit.xSwitch_CoolWind;
i_pstStSysParam^.astStRSV_UnitParam_Save[iUnitId].byGetErrMode:=
			i_pstStParam_Diamonds_WrRd^.astStWrRd_UnitParam[iUnitId].byGetErrMode;
END_FOR
//在这里处理一下减速比单独设定和周长单独设定问题；
i_pstStSysParam^.stStSysParam_Save.wCtlFlag_IndependentSettings.0:= i_pstStParam_Diamonds_WrRd^.stBitStWrRd_Switch_Machine.xSwitch_IndependentSettings_BottomGirth;
i_pstStSysParam^.stStSysParam_Save.wCtlFlag_IndependentSettings.2:= i_pstStParam_Diamonds_WrRd^.stBitStWrRd_Switch_Machine.xSwitch_IndependentSettings_NetGirth;
i_pstStSysParam^.stStSysParam_Save.wCtlFlag_IndependentSettings.8:= i_pstStParam_Diamonds_WrRd^.stBitStWrRd_Switch_Machine.xSwitch_IndependentSettings_BottomRatio;
i_pstStSysParam^.stStSysParam_Save.wCtlFlag_IndependentSettings.10:= i_pstStParam_Diamonds_WrRd^.stBitStWrRd_Switch_Machine.xSwitch_IndependentSettings_NetRatio;

IF i_pstStParam_Diamonds_WrRd^.stBitStWrRd_Switch_Machine.xSwitch_IndependentSettings_BottomGirth THEN//底辊周长单独设定
	//这时候只更新色组底辊周长
	FOR iUnitId:=1 TO MAX_UNIT_NUM BY 1 DO
		i_pstStSysParam^.astStUnitParam_Save[iUnitId].rGirth_BottomRoller:= i_pstStParam_Diamonds_WrRd^.astStWrRd_UnitParam[iUnitId].rGirth_BottomGirth;
	END_FOR
ELSE
	FOR iGrp:=1 TO 2 BY 1 DO
		i_pstStSysParam^.astStGrpParam_Save[iGrp].rGirth_BottomRoller:= i_pstStParam_Diamonds_WrRd^.arGirth_BottomRoller[iGrp];
	END_FOR
END_IF
IF i_pstStParam_Diamonds_WrRd^.stBitStWrRd_Switch_Machine.xSwitch_IndependentSettings_NetGirth THEN//底辊周长单独设定
	//这时候只更新色组wang辊周长
	FOR iUnitId:=1 TO MAX_UNIT_NUM BY 1 DO
		i_pstStSysParam^.astStUnitParam_Save[iUnitId].rGirth_NetRoller:= i_pstStParam_Diamonds_WrRd^.astStWrRd_UnitParam[iUnitId].rGirth_NetGirth;
	END_FOR
ELSE
	FOR iGrp:=1 TO 2 BY 1 DO
		i_pstStSysParam^.astStGrpParam_Save[iGrp].rGirth_NetRoller:= i_pstStParam_Diamonds_WrRd^.arGirth_NetRoller[iGrp];
	END_FOR
END_IF
//底辊减速比
IF i_pstStParam_Diamonds_WrRd^.stBitStWrRd_Switch_Machine.xSwitch_IndependentSettings_BottomRatio THEN//底辊周长单独设定
	//这时候只更新色组wang辊周长
	FOR iUnitId:=1 TO MAX_UNIT_NUM BY 1 DO
		i_pstStSysParam^.astStUnitParam_Save[iUnitId].uiNum_BottomRoller:= i_pstStParam_Diamonds_WrRd^.astStWrRd_UnitParam[iUnitId].uiNum_Bottom;
		i_pstStSysParam^.astStUnitParam_Save[iUnitId].uiDen_BottomRoller:= i_pstStParam_Diamonds_WrRd^.astStWrRd_UnitParam[iUnitId].uiDen_Bottom;
	END_FOR
ELSE
	FOR iGrp:=1 TO 2 BY 1 DO
		i_pstStSysParam^.astStGrpParam_Save[iGrp].uiNum_BottomRoller:= i_pstStParam_Diamonds_WrRd^.auiNum_BottomRoller[iGrp];
		i_pstStSysParam^.astStGrpParam_Save[iGrp].uiDen_BottomRoller:= i_pstStParam_Diamonds_WrRd^.auiDen_BottomRoller[iGrp];
	END_FOR
END_IF
//wang辊减速比
IF i_pstStParam_Diamonds_WrRd^.stBitStWrRd_Switch_Machine.xSwitch_IndependentSettings_NetRatio THEN//底辊周长单独设定
	//这时候只更新色组wang辊周长
	FOR iUnitId:=1 TO MAX_UNIT_NUM BY 1 DO
		i_pstStSysParam^.astStUnitParam_Save[iUnitId].uiNum_NetRoller:= i_pstStParam_Diamonds_WrRd^.astStWrRd_UnitParam[iUnitId].uiNum_Net;
		i_pstStSysParam^.astStUnitParam_Save[iUnitId].uiDen_NetRoller:= i_pstStParam_Diamonds_WrRd^.astStWrRd_UnitParam[iUnitId].uiDen_Net;
	END_FOR
ELSE
	FOR iGrp:=1 TO 2 BY 1 DO
		i_pstStSysParam^.astStGrpParam_Save[iGrp].uiNum_NetRoller:= i_pstStParam_Diamonds_WrRd^.auiNum_NetRoller[iGrp];
		i_pstStSysParam^.astStGrpParam_Save[iGrp].uiDen_NetRoller:= i_pstStParam_Diamonds_WrRd^.auiDen_NetRoller[iGrp];
	END_FOR
END_IF

i_pstStSysParam^.astStUnitParam_Save[1].iMarkArrangeMode;
i_pstStSysParam^.astStUnitParam_Save[2].iMarkArrangeMode;
i_pstStSysParam^.astStUnitParam_Save[3].iMarkArrangeMode;
i_pstStSysParam^.astStUnitParam_Save[4].iMarkArrangeMode;
i_pstStSysParam^.astStUnitParam_Save[5].iMarkArrangeMode;
i_pstStSysParam^.astStUnitParam_Save[6].iMarkArrangeMode;
i_pstStSysParam^.astStUnitParam_Save[7].iMarkArrangeMode;
i_pstStSysParam^.astStUnitParam_Save[8].iMarkArrangeMode;
i_pstStSysParam^.astStUnitParam_Save[9].iMarkArrangeMode;
i_pstStParam_Diamonds_WrRd^.astStWrRd_UnitParam[1].iMarkArrangeMode;
i_pstStParam_Diamonds_WrRd^.astStWrRd_UnitParam[2].iMarkArrangeMode;
i_pstStParam_Diamonds_WrRd^.astStWrRd_UnitParam[3].iMarkArrangeMode;
i_pstStParam_Diamonds_WrRd^.astStWrRd_UnitParam[4].iMarkArrangeMode;
i_pstStParam_Diamonds_WrRd^.astStWrRd_UnitParam[5].iMarkArrangeMode;
i_pstStParam_Diamonds_WrRd^.astStWrRd_UnitParam[6].iMarkArrangeMode;
i_pstStParam_Diamonds_WrRd^.astStWrRd_UnitParam[7].iMarkArrangeMode;
i_pstStParam_Diamonds_WrRd^.astStWrRd_UnitParam[8].iMarkArrangeMode;
i_pstStParam_Diamonds_WrRd^.astStWrRd_UnitParam[9].iMarkArrangeMode;
(*2025.10.23.135406*)
Action_Output_SysCfg_Rd();

//2025.10.22.091027 | bai.zy | 配方

//2025.10.22.091027 | bai.zy | 配方
FOR iGrp := 1 TO 2 BY 1 DO
	//获取启动标志@2026.5.24.212821+
	afbRestorePhase[iGrp](CLK:=i_pstStParam_Diamonds_WrRd^.astBitStWrRd_Switch_Grp[iGrp].xBtn_RestorePhase_Hmi);
	i_pstStParam_Diamonds_WrRd^.astBitStWrRd_Switch_Grp[iGrp].xBtn_RestorePhase_Hmi:= FALSE;
	IF afbRestorePhase[iGrp].Q THEN

		ax_RestorePhase_hmi[iGrp] := TRUE;
	END_IF

	IF ax_RestorePhase_hmi[iGrp] THEN
		//2026.5.15.113637校验
		IF NOT axInitTime[iGrp] THEN

			tmStart_ReadPhase:= TIME();
			axInitTime[iGrp]:= TRUE;
			g_axPhaseRestore_Overtime[iGrp] := FALSE;

		END_IF

		wChk_Tmp:= KS_CRC(i_pstStRd_PhaseRead,SIZEOF(i_pstStRd_PhaseRead^)-6,ADR(dwSum_Tmp));
		IF TIME()-tmStart_ReadPhase<tmTimeOut_ReadPhase THEN//判断超时时间
			IF wChk_Tmp= i_pstStRd_PhaseRead^.wChk AND
					dwSum_Tmp= i_pstStRd_PhaseRead^.dwSum AND
					dwSum_Tmp<> 0 THEN

				i_pstStSysParam^.astStGrpParam_Save[iGrp].rGirth_PrnRoller 	:= i_pstStRd_PhaseRead^.arGirth_Pu[iGrp];
				i_pstStSysParam^.astStGrpParam_Save[iGrp].iMarkTypeId 		:= i_pstStRd_PhaseRead^.aiMarkTypeId[iGrp];
				i_pstStSysParam^.astStGrpParam_Save[iGrp].iMarkArrangeMode  := i_pstStRd_PhaseRead^.aiMarkArrangeId[iGrp];
				i_pstStSysParam^.astStGrpParam_Save[iGrp].byTriMark_SideC   := i_pstStRd_PhaseRead^.abyTriMark_SideC[iGrp];
				i_pstStSysParam^.astStGrpParam_Save[iGrp].byTriMark_SideB   := i_pstStRd_PhaseRead^.abyTriMark_SideB[iGrp];
				//是不是和下面这个变量是一样的作用？？？
				//i_pstStSysParam^.stStSysParam_Save.wCtlFlag_IndependentSettings.1 := i_pstStRd_PhaseRead^.axGirthInputMode[iGrp];

				i_pstStSysParam^.astStGrpParam_Save[iGrp].rTaper_Begin_If   := i_pstStRd_PhaseRead^.arTaper_Begin_If[iGrp];
				i_pstStSysParam^.astStGrpParam_Save[iGrp].rTaper_End_If     := i_pstStRd_PhaseRead^.arTaper_End_If[iGrp];
				i_pstStSysParam^.astStGrpParam_Save[iGrp].rTaper_Begin_Of   := i_pstStRd_PhaseRead^.arTaper_Begin_Of[iGrp];
				i_pstStSysParam^.astStGrpParam_Save[iGrp].rTaper_End_Of     := i_pstStRd_PhaseRead^.arTaper_End_Of[iGrp];
				i_pstStSysParam^.astStGrpParam_Save[iGrp].rTaper_Begin_Uw   := i_pstStRd_PhaseRead^.arTaper_Begin_Uw[iGrp];
				i_pstStSysParam^.astStGrpParam_Save[iGrp].rTaper_End_Uw     := i_pstStRd_PhaseRead^.arTaper_End_Uw[iGrp];
				i_pstStSysParam^.astStGrpParam_Save[iGrp].rTaper_Begin_Rw   := i_pstStRd_PhaseRead^.arTaper_Begin_Rw[iGrp];
				i_pstStSysParam^.astStGrpParam_Save[iGrp].rTaper_End_Rw     := i_pstStRd_PhaseRead^.arTaper_End_Rw[iGrp];

				FOR iUnitId := 1 TO MAX_UNIT_NUM BY 1 DO
					i_pstStSysParam^.astStUnitParam_Save[iUnitId].rGirth_PrnRoller 					:= i_pstStRd_PhaseRead^.arGirth[iUnitId];
					i_pstStSysParam^.astStUnitParam_Save[iUnitId].xEnable_Arc                       := i_pstStRd_PhaseRead^.axEnable_Arc[iUnitId];
					i_pstStSysParam^.astStUnitParam_Save[iUnitId].iMarkTypeId                       := i_pstStRd_PhaseRead^.aiMarkTypeId_Pu[iUnitId];
					i_pstStSysParam^.astStUnitParam_Save[iUnitId].iMarkArrangeMode                  := i_pstStRd_PhaseRead^.aiMarkArrangeId_Pu[iUnitId];
					i_pstStSysParam^.astStUnitParam_Save[iUnitId].iGateWidthPhy                     := i_pstStRd_PhaseRead^.aiGateWidthPhy[iUnitId];
					i_pstStSysParam^.astStUnitParam_Save[iUnitId].iGateSa                           := i_pstStRd_PhaseRead^.aiGateSa[iUnitId];
					i_pstStSysParam^.astStUnitParam_Save[iUnitId].iGateSaEx                         := i_pstStRd_PhaseRead^.aiGateSaEx[iUnitId];
					i_pstStSysParam^.astStUnitParam_Save[iUnitId].dwFlag_Ctl.0 := i_pstStRd_PhaseRead^.abySwitch_Unit_Phase[iUnitId].0;
					i_pstStSysParam^.astStUnitParam_Save[iUnitId].dwFlag_Ctl.2 := i_pstStRd_PhaseRead^.abySwitch_Unit_Phase[iUnitId].1;
					i_pstStSysParam^.astStUnitParam_Save[iUnitId].dwFlag_Ctl.3 := i_pstStRd_PhaseRead^.abySwitch_Unit_Phase[iUnitId].2;
					i_pstStSysParam^.astStUnitParam_Save[iUnitId].dwFlag_Ctl.11 := i_pstStRd_PhaseRead^.abySwitch_Unit_Phase[iUnitId].3;
					i_pstStSysParam^.astStUnitParam_Save[iUnitId].dwFlag_Ctl.12 := i_pstStRd_PhaseRead^.abySwitch_Unit_Phase[iUnitId].4;
					i_pstStSysParam^.astStUnitParam_Save[iUnitId].xSwitchOn_CoatingPrn := i_pstStRd_PhaseRead^.abySwitch_Unit_Phase[iUnitId].5;
					i_pstStSysParam^.astStUnitParam_Save[iUnitId].rAdj_V                            := i_pstStRd_PhaseRead^.arAdj_V[iUnitId];
					i_pstStSysParam^.astStUnitParam_Save[iUnitId].rAdj_H                            := i_pstStRd_PhaseRead^.arAdj_H[iUnitId];
					i_pstStSysParam^.astStUnitParam_Save[iUnitId].iPhase_RegisterOK                 := i_pstStRd_PhaseRead^.aiPhase_RegisterOK[iUnitId];
					i_pstStSysParam^.astStUnitParam_Save[iUnitId].rSV_UnitTemCtl                    := i_pstStRd_PhaseRead^.arSV_TemCtl[iUnitId];
					i_pstStSysParam^.astStUnitParam_Save[iUnitId].byHotBlower_AO          			:= i_pstStRd_PhaseRead^.abyAiirInletWindDoorValue[iUnitId];
					i_pstStSysParam^.astStUnitParam_Save[iUnitId].byOvensAirOutWindDoorValue        := i_pstStRd_PhaseRead^.abyOvensAirOutWindDoorValue[iUnitId];
					i_pstStSysParam^.astStUnitParam_Save[iUnitId].wAirExhaustWindDoorValue         	:= i_pstStRd_PhaseRead^.abyAirExhaustWindDoorValue[iUnitId];
					i_pstStSysParam^.astStUnitParam_Save[iUnitId].wAirReturnWindDoorValue          	:= i_pstStRd_PhaseRead^.abyAirReturnWindDoorValue[iUnitId];
					i_pstStSysParam^.astStUnitParam_Save[iUnitId].rHz_UnitInkRoller_ManuallySet     := i_pstStRd_PhaseRead^.arHz_UnitInkRoller_ManuallySet[iUnitId];
					i_pstStSysParam^.astStUnitParam_Save[iUnitId].rCoeff_UnitInkRoller_Auto         := i_pstStRd_PhaseRead^.arCoeff_UnitInkRoller_Auto[iUnitId];
					i_pstStSysParam^.astStUnitParam_Save[iUnitId].rHz_UnitScraper_ManuallySet       := i_pstStRd_PhaseRead^.arHz_UnitScraper_ManuallySet[iUnitId];
					i_pstStSysParam^.astStUnitParam_Save[iUnitId].rCoeff_UnitScraper_Auto           := i_pstStRd_PhaseRead^.arCoeff_UnitScraper_Auto[iUnitId];
					i_pstStSysParam^.astStUnitParam_Save[iUnitId].rHz_UnitHotWind_ManuallySet       := i_pstStRd_PhaseRead^.arHz_UnitHotWind_ManuallySet[iUnitId];
					i_pstStSysParam^.astStUnitParam_Save[iUnitId].rHz_UnitHotWind_2_ManuallySet     := i_pstStRd_PhaseRead^.arHz_UnitHotWind_2_ManuallySet[iUnitId];
					i_pstStSysParam^.astStUnitParam_Save[iUnitId].rHz_UnitExhaust_ManuallySet       := i_pstStRd_PhaseRead^.arHz_UnitExhaust_ManuallySet[iUnitId];
				END_FOR

				i_pstStSysParam^.astStGrpParam_UnSave[iGrp].xFlag_PhaseRestore := TRUE;
				axInitTime[iGrp]:= FALSE;

				//这里只先清空一下校验码吧
				i_pstStRd_PhaseRead^.wChk:= 0;
				i_pstStRd_PhaseRead^.dwSum:= 0;
				ax_RestorePhase_hmi[iGrp]:= FALSE;
			END_IF
		ELSE
			axInitTime[iGrp]:= FALSE;

			i_pstStSysParam^.astStGrpParam_UnSave[iGrp].xFlag_PhaseRestore := FALSE;
			//增加一个报警码？
			//报警清除在Action_Alarm_ClearAndReset，直接清除这个标志
			g_axPhaseRestore_Overtime[iGrp] := TRUE;

			ax_RestorePhase_hmi[iGrp]:= FALSE;//超时直接处理清除
		END_IF

	END_IF

// 	//恢复相位完成了也清除一次
// 	afbResetRestorePhase[iGrp](CLK:= NOT i_pstStSysParam^.astStGrpParam_UnSave[iGrp].xFlag_PhaseRestore);
// 	//IF afbResetRestorePhase[iGrp].Q THEN

// 	IF (NOT i_pstStSysParam^.astStGrpParam_UnSave[iGrp].xFlag_PhaseRestore) AND
// 		(NOT i_pstStParam_Diamonds_WrRd^.astBitStWrRd_Switch_Grp[iGrp].xBtn_RestorePhase_Hmi) THEN
// // 		xInitTime:= FALSE;
// 		ax_RestorePhase_hmi[iGrp]:= FALSE;//超时直接处理清除
// 	END_IF
	(**)

	//读取装版相位
	IF  i_pstStParam_Diamonds_WrRd^.astBitStWrRd_Switch_Grp[iGrp].xBtn_ReadPhase_Home THEN
		i_pstStParam_Diamonds_WrRd^.astBitStWrRd_Switch_Grp[iGrp].xBtn_ReadPhase_Home := FALSE;
		i_pstStSysParam^.astStGrpParam_UnSave[iGrp].xBtn_Home := TRUE;
	END_IF

		//2026.1.26.171345 | + | 增加回零位的功能
	IF g_axBackToHome[iGrp] OR i_pstStParam_Diamonds_WrRd^.astBitStWrRd_Switch_Grp[iGrp].xSwitch_BackToHome THEN
		g_axBackToHome[iGrp] := FALSE;
		i_pstStParam_Diamonds_WrRd^.astBitStWrRd_Switch_Grp[iGrp].xSwitch_BackToHome := FALSE;
		i_pstStSysParam^.astStGrpParam_UnSave[iGrp].xFlag_PhaseRestore := TRUE;
		FOR iUnitId := 1 TO MAX_UNIT_NUM BY 1 DO
			i_pstStSysParam^.astStUnitParam_Save[iUnitId].iPhase_RegisterOK := 0;
		END_FOR
	END_IF

END_FOR
